(* IEC 61131-3 sources: plcassist-cli/packages/volt-lsp-iec/test-corpus/pro2193/Device/Plc Logic/Application/09 Misc/Library Manager/L_MC1P_MotionControlBasic (part 2) *)

(* ---- AXIS_REF.fb ---- *)
FUNCTION_BLOCK AXIS_REF EXTENDS L_DCO_AXIS_REF_BASE
VAR_INPUT
	LRVELOVERRIDE : LREAL := 1.0;
	LRACCOVERRIDE : LREAL := 1.0;
	LRJERKOVERRIDE : LREAL := 1.0;
	LRCOMMANDEDPOSITION : LREAL;
	LRCOMMANDEDVELOCITY : LREAL;
	LRCOMMANDEDACCELERATION : LREAL;
	LRSETVELOCITYLIMITHIGH : LREAL := 0;
	LRSETVELOCITYLIMITLOW : LREAL := 0;
	LRTORQUELIMHIGH : LREAL;
	LRTORQUELIMLOW : LREAL;
	LRTORQUELIMAUX : LREAL;
	SITORQUELIMDIR : SINT;
	XDELETETORQUELIM : BOOL;
	XSETTORQUELIMAUX : BOOL;
	XTORQUELIMHIGHFROMAPP : BOOL;
	XTORQUELIMLOWFROMAPP : BOOL;
	ITORQUELIMHIGHPCT : INT := 2000;
	ITORQUELIMLOWPCT : INT := 2000;
	EDIRECTION : MC_DIRECTION;
	XDRIVEENABLE : BOOL;
	XERRORRESET : BOOL;
	LRREFOFFSET : LREAL;
	LRREFOFFSETACT : LREAL;
	XENABLEPOSITIVE : BOOL := TRUE;
	XENABLENEGATIVE : BOOL := TRUE;
	LRSETSUPERACC : LREAL;
	LRSETSUPERVEL : LREAL;
	LRSETSUPERPOS : LREAL;
	LRSETMOVEACC : LREAL;
	LRSETMOVEVEL : LREAL;
	LRSETMOVEPOS : LREAL;
	XBUFCMDDONE : BOOL;
	XBUFRESTART : BOOL;
	LRPROFILESPEEDFIRST : LREAL;
	LRPROFILETARGETSPEED : LREAL;
	DWBUFFERCMD : __XWORD;
	XDISABLEERRORLOGGING : BOOL;
	XMOVEFUNBUSY : BOOL;
	XSUPERFUNBUSY : BOOL;
	LRCOMMANDEDPOSABSOLUT : LREAL;
	XRESETFOLLOWINGERROR : BOOL;
	XSETAXISQSP : BOOL;
	XSETDRIVEQSP : BOOL;
	EAXISSTATE : L_MC1P_AXIS_STATE := 2;
	LRSETPOSITION : LREAL := 0.0;
	LRSETVELOCITY : LREAL := 0.0;
	LRSETACCELERATION : LREAL := 0.0;
	LRSETTORQUE : LREAL := 0.0;
	LRVLTARGETVEL : LREAL := 0.0;
	LRLIMITEDVELOCITY : ARRAY [1..4] OF LREAL;
	LRLIMITEDDECTIME : ARRAY [1..4] OF LREAL;
	LRRESETSLSOFFSETVELOCITY : LREAL;
	DWLIMITERCONTROLACT : DWORD;
	SCSTOPAXISBYAPPL : L_MC1P_StopOperation;
	XSTAYINLASTSTATEREQUEST : BOOL;
	XMOVELASTSETPOSREQUEST : BOOL;
	LRSETVELMOVELASTSETPOS : LREAL;
	LRSETACCMOVELASTSETPOS : LREAL;
	LRSETDECMOVELASTSETPOS : LREAL;
	LRSETJERKMOVELASTSETPOS : LREAL;
	EDIRECTIONMOVELASTSETPOS : MC_DIRECTION;
	EDIRECTIONACTPROFILE : MC_DIRECTION;
	WAXISCONTROL : WORD := 0;
	XALLOWCHANGEOFCINHPAR : BOOL := FALSE;
	LRMOVEVELOFFSETVEL : LREAL;
	EOPTIMIZEDPROFILECALCULATIONMODE : UINT := 1;
	XLEAVESERVICESTATE : BOOL;
	XLEAVESERVICESTATEDISABLEDRIVE : BOOL;
	WLEAVESERVICESTATEPOWID : WORD;
END_VAR
VAR_OUTPUT
	EDEVICE : L_MC1P_DriveType := 0;
	WAXISSTATUS : DWORD := 0;
	EACTIVEERRORID : WORD := 0;
	LRACTPOSITION : LREAL := 0.0;
	LRACTVELOCITY : LREAL := 0.0;
	LRACTACCELERATION : LREAL := 0.0;
	LRACTTORQUE : LREAL := 0.0;
	LRSETTORQUETODRIVE : LREAL := 0;
	LRACTFOLLOWINGERROR : LREAL := 0.0;
	LRMAXFOLLOWINGERROR : LREAL := 0.0;
	XVIRTUAL : BOOL;
	XAXISAVAILABLE : BOOL;
	EACTDIRECTION : MC_DIRECTION;
	LRDIRECTIONHYSTERESISPOS : LREAL;
	LRDIRECTIONHYSTERESISTOL : LREAL := 1E-06;
	XDRIVEENABLED : BOOL;
	XERROR : BOOL;
	XWARNING : BOOL;
	XDRIVEERROR : BOOL;
	XDRIVEWARNING : BOOL;
	DWDRIVEERRORID : DWORD;
	XHOMEPOSAVAILABLE : BOOL;
	XSWLIMITENABLED : BOOL;
	XSWLIMITPOS : BOOL;
	XSWLIMITNEG : BOOL;
	XHWLIMITPOS : BOOL;
	XHWLIMITNEG : BOOL;
	XSPEEDEQZERO : BOOL;
	XINPOSITION : BOOL;
	LRTASKCYCLE : LREAL := 0.001;
	LRINVTASKCYCLE : LREAL := 1000.0;
	LRSWLIMITPOS : LREAL := 0.0;
	LRSWLIMITNEG : LREAL := 0.0;
	LRLASTSETPOSITION : LREAL;
	LRLASTTARGETPOSITION : LREAL;
	XSTANDSTILLSETVELOCITY : BOOL;
	XSTANDSTILLACTVELOCITY : BOOL;
	XSTOACTIVE : BOOL;
	XVOLTAGEENABLED : BOOL;
	XAXISREADYTOSWITCHON : BOOL;
	XAXISREADYFORMOTION : BOOL;
	SCPAR : L_MC1P_ParAccess;
END_VAR
VAR
	DWAXISCONFIGSETTINGS : DWORD;
	XSETVALUESAVAILABLE : BOOL;
	BYSETVALUESVALID : BYTE;
	DWTASKYCLE_US : DWORD := 1000;
	XSUSPENDFOLLOWINGERRORINT : BOOL;
	XSUSPENDFOLLOWINGERROREXT : BOOL;
	LRMAXVELOCITYAPPLOLD : LREAL;
	LRMAXACCELERATIONAPPLOLD : LREAL;
	LRMAXJERKAPPLOLD : LREAL;
	LRSWLIMITPOSOLD : LREAL;
	LRSWLIMITNEGOLD : LREAL;
	XENABLEPOSOLD : BOOL;
	XENABLENEGOLD : BOOL;
	DWLIMITERCONTROLOLD : DWORD;
	LRLIMITEDVELOCITYOLD : ARRAY [1..4] OF LREAL;
	LRLIMITEDDECTIMEOLD : ARRAY [1..4] OF LREAL;
	LRLIMITEDJERKOLD : ARRAY [1..4] OF LREAL;
	ELIMITERSTOPREACTION : L_IE1P_SeverityLevel := L_IE1P_SeverityLevel.WARNING;
	XSWLIMITDISABLE : BOOL := FALSE;
	XSWLIMITPOSNEU : BOOL;
	XSWLIMITPOSISTAN : BOOL;
	XSWLIMITNEGNEU : BOOL;
	XSWLIMITNEGISTAN : BOOL;
	PBYCOUPLEDMASTERAXIS : POINTER TO BYTE;
	PBYCOUPLEDPHASINGMASTERAXIS : POINTER TO BYTE;
	LRPHASESHIFTPOS : LREAL;
	LRPHASESHIFTVEL : LREAL;
	LRPHASESHIFTACC : LREAL;
	LRPHASESHIFTPOSOLD : LREAL;
	LRPHASESHIFTVELOLD : LREAL;
	LRPHASESHIFTACCOLD : LREAL;
	XSETPHASESHIFTVALUES : BOOL;
	ETRAVERSINGRANGEACT : L_MC1P_TraversingRange := 0;
	LRCYCLELENGTHACT : LREAL := 360.0;
	XENABLEHWLIMITPOS : BOOL := TRUE;
	XENABLEHWLIMITNEG : BOOL := TRUE;
	XHWSIGNALNEG : BOOL := FALSE;
	XHWSIGNALPOS : BOOL := FALSE;
	BHWENSCHPOSNEU : BOOL := TRUE;
	BNOTIFYERRORHWLIMITPOSISTAN : BOOL;
	BHWENSCHNEGNEU : BOOL := TRUE;
	BNOTIFYERRORHWLIMITNEGISTAN : BOOL;
	XAXISISHOMESOURCE : BOOL;
	XHOMEPOSAVAILABLEDRIVE : BOOL;
	SCHOMEPARAMETER : L_MC1P_HomeParameter;
	LRHOMEPOSITION : LREAL;
	XPOSCTRL : BOOL;
	XTPSUPPORTED : BOOL := FALSE;
	XTPWITHTIMESTAMP : BOOL := FALSE;
	SNTPMAXCHANNEL : SINT;
	PG : L_MC1P_PosProfiler := STRUCT(wCalcProfileMode := 1);
	ITFPG_MOVEACTIVE : L_MC1P_IPosProfilerActive;
	PG_MOVE : L_MC1P_PosProfiler := STRUCT(wCalcProfileMode := 1);
	ITFPG_SUPERACTIVE : L_MC1P_IPosProfilerActive;
	PG_SUPER : L_MC1P_PosProfiler := STRUCT(wCalcProfileMode := 1);
	PG_DUMMY : L_MC1P_PosProfiler := STRUCT(wCalcProfileMode := 1);
	SCPARAMSTOP : L_MC1P_ProfileParameter;
	XCTRLMODECHANGEREQ : BOOL;
	LRCTRLMODECHANGEREQACTVEL : LREAL;
	PFBMOVEBASIC : POINTER TO L_MC1P_MoveBasic;
	PFBMOVEBASICSUPER : POINTER TO L_MC1P_MoveBasic;
	XRESTARTPOSITIONING : BOOL;
	LRSETPOSITIONOLD : LREAL;
	LRSETVELOCITYOLD : LREAL;
	LRSETACCELERATIONOLD : LREAL;
	WACTFUNID : WORD := 0;
	WACTSUPERFUNID : WORD := 0;
	WACTPHASEFUNID : WORD := 0;
	PSERRORINST : POINTER TO STRING;
	SERRORINST : STRING;
	ERRORMANAGER : L_IE1P_ErrorManager;
	ERRORRESETOCCUREDTIMEWITHOUTLEM : SYSTIME;
	ASCERRORINFO : REFERENCE TO ARRAY [0..7] OF L_IE1P_ErrorInformation;
	ASCWARNINGINFO : REFERENCE TO ARRAY [0..7] OF L_IE1P_ErrorInformation;
	WINITSTATE : WORD;
	PAPPLICATION : POINTER TO APPLICATION;
	ATPDATA : ARRAY [1..4] OF L_MC1P_TPData;
	ATPDATASAVE : L_MC1P_TPData;
	XHOMINGSUPPORTED : BOOL;
	EAXISSTATEOLD : L_MC1P_AXIS_STATE := L_MC1P_AXIS_STATE.Disabled;
	ECONTROLMODE : L_MC1P_ControlMode := L_MC1P_ControlMode.PosCtrlDrive;
	ECONTROLMODEDEFAULT : L_MC1P_ControlMode := L_MC1P_ControlMode.PosCtrlDrive;
	ECONTROLMODEDEFAULTINT : L_MC1P_ControlMode := L_MC1P_ControlMode.PosCtrlDrive;
	POSCTRLDRIVEAVAILABLE : L_IE1P_Error;
	POSCTRLPLCAVAILABLE : L_IE1P_Error;
	SPEEDCTRLDRIVEAVAILABLE : L_IE1P_Error;
	TORQUECTRLDRIVE : L_IE1P_Error;
	XDRIVEENABLEOLD : BOOL;
	XLOCKEDFORSINGLEMOTION : BOOL := FALSE;
	XHOMEABSSWITCH : BOOL;
	XHOMEABSSWITCHOVERWRITEACTIVE : BOOL;
	XRAMPTOSTANDSTILL : BOOL;
	XRAMPTOSTANDSTILLDONE : BOOL;
	XRAMPTOSTANDSTILLACTIVE : BOOL;
	XDRIVEENABLEDOLD : BOOL;
	XDRIVEENABLEDREAL : BOOL;
	XDRIVEENABLEDREALOLD : BOOL;
	LRFOLLOWINGERRORINT : LREAL;
	XSUPPORTBRAKE : BOOL := FALSE;
	XSUPPORTDCBRAKE : BOOL := FALSE;
	XUSEASVIRTUALEXT : BOOL := FALSE;
	XUSEASVIRTUALEXTACT : BOOL := FALSE;
	LRSETSUPERACCOLD : LREAL;
	LRSETSUPERVELOLD : LREAL;
	LRSETSUPERPOSOLD : LREAL;
	ITFPARA : L_MC1P_IPara;
	XFASTSTOPDONE : BOOL;
	XFASTSTOPDONESAVE : BOOL;
	XSETFASTSTOPINT : BOOL;
	XERRRORSTOPACTIVE : BOOL;
	XERRRORSTOPDONE : BOOL;
	XSETAXISQSPACTIVE : BOOL;
	XRAMPQSPSTARTCALLEDFROMAPP : BOOL;
	XDRIVEQSPACTIVE : BOOL;
	XDRIVEQSPACTIVEOLD : BOOL;
	XDRIVEQSPSET : BOOL;
	XSETDRIVEFAILQSP : BOOL;
	XSETDRIVEFAILCINH : BOOL;
	XDRIVEQSPDONE : BOOL;
	XDRIVEQSPDONESAVE : BOOL;
	ESTOPTYPE : WORD;
	POW : L_MC1P_Power_Internal;
	XOBERVERESWITCHONTIME : BOOL := TRUE;
	FBBASE : L_MC1P_Template_ForAxis;
	ABC : L_MC1P_AxisBasicControl_Internal;
	ABCDATA : L_MC1P_AxisBasicControlInstanceData;
	ITFENCODER : L_MC1P_IEncoderInterface;
	ITFENCODERHANDLER : L_MC1P_IEncoderInterface;
	LRSETTORQUEFROMAXESGROUP : LREAL := 0;
	EPRECONTROLMODE : L_MC1P_PreControlMode := L_MC1P_PreControlMode.Automatic;
	GUID : L_MC1P_AxisGUID;
	LRTORQUEPRECTRL : LREAL;
	LRTORQUESET : LREAL;
	XMOVEFUNBUSYOLD : BOOL;
	XMOVEFUNBUSYOLDOLD : BOOL;
	DWIODRVDEVICEID : DWORD;
	WIODRVDEVICETYPE : WORD;
	EDEVICEORIGIN : L_MC1P_DriveType := L_MC1P_DriveType.Virtual;
	EDEVICECLASS : L_MC1P_DeviceClass := L_MC1P_DeviceClass.VirtualAxis;
	DWTARGETID : DWORD := 0;
	XCTRLFIRMWARECHECKPASSED : BOOL := FALSE;
	XENABLELOGENTRY : BOOL := 1;
	ETRAVERSINGRANGE : L_MC1P_TraversingRange := 1;
	LRCYCLELENGTH : LREAL := 360.0;
	LRINVCYCLELENGTH : LREAL := (1.0 / 360.0);
	LRDEFAULTVELOCITY : LREAL := 0.0;
	LRDEFAULTACCELERATION : LREAL := 0.0;
	LRDEFAULTJERK : LREAL := 0.0;
	LRMAXVELOCITYAPPL : LREAL := 0.0;
	LRMAXACCELERATIONAPPL : LREAL := 0.0;
	LRMAXJERKAPPL : LREAL := 0.0;
	XENABLESWLIMIT : BOOL := 0;
	WBEHAVEONSWLIMIT : WORD := 1;
	LRDECERRORSTOP : LREAL := 3600.0;
	LRJERKERRORSTOP : LREAL := 0.0;
	XREAKTONMCFBERROR : BOOL := 1;
	LRWINDOWSTANDSTILL : LREAL := 0.0;
	LRWINDOWVELOCITYCONST : LREAL := 0.0;
	LRWINDOWTARGETREACHED : LREAL := 0.0;
	LRWINDOWTARGETREACHEDTIME : LREAL := 0.0;
	LRMODPOSTOLERANCE : LREAL := 0.0;
	XSETVALUEMONITORING : BOOL := 0;
	EPARAMETERINDEX : WORD := 101;
	DWPARABASEINDEX : DWORD;
	PPARA2 : L_SSYP.L_SSYP_EVTPARAM_CmpLenzeIPCSystemSoftPLCParaChanged;
	HEVENTPARWRITE : SysTypes.RTS_IEC_HANDLE;
	HINTERFACEPARWRITE : SysTypes.RTS_IEC_HANDLE;
	HEVENTDOWNLOADDONE : SysTypes.RTS_IEC_HANDLE;
	HINTERFACEDOWNLOADDONE : SysTypes.RTS_IEC_HANDLE;
	HEVENTRESETDONE : SysTypes.RTS_IEC_HANDLE;
	HINTERFACERESETDONE : SysTypes.RTS_IEC_HANDLE;
	ITFCALLBACK : CmpEventMgr.ICmpEventCallback;
	DWEVENTCOUNTER : DWORD;
	WENABLEDRIVEBLOCKEDBYOBJECTTRANSFER : WORD := 0;
	XUSEDBYAXESGROUP : BOOL;
	PUSEDAXESGROUP : POINTER TO BYTE;
	DWEVTINITCOUNT : DWORD;
	XNEWHOMEPOSLOADED : BOOL;
	DWSETPOSITIONCALLCYCLE : DWORD;
	XSETPOSITIONCALLCYCLEVALID : BOOL;
	AITFFILTER : ARRAY [1..c_MaxFilterInt] OF L_MC1P_ISetvalueManipulationInterface;
	XENABLEFILTER : BOOL;
	XFILTERAVAILABLE : BOOL;
	XIGNORFILTERINSTOP : BOOL := TRUE;
	XIGNORFILTERINSTOPITF : BOOL;
	XUSEFILTERVALUESFORSYNC : BOOL := FALSE;
	LRSETPOSITIONFILT : LREAL;
	LRSETVELOCITYFILT : LREAL;
	LRSETACCELERATIONFILT : LREAL;
	LRSETTORQUEFILT : LREAL;
	LRSETVALUEFILTERPOSDEVIATION : LREAL;
	XINTARGETSETVALUEFILTER : BOOL;
	XSUSPENDSETVALUEFILTERCALL : BOOL := FALSE;
	LRSETPOSITIONFILTOLD : LREAL;
	LRSETVELOCITYFILTOLD : LREAL;
	LRSETACCELERATIONFILTOLD : LREAL;
	LRSETTORQUEFILTOLD : LREAL;
	LRSETPOSROUNDSFILTOLD : LREAL;
	AITFCOMPENSATION : ARRAY [1..c_MaxFilterInt] OF L_MC1P_ICompensationInterface;
	LRCOMPENSATIONOFFSETPOS : LREAL;
	LRCOMPENSATIONOFFSETVEL : LREAL;
	LRCOMPENSATIONOFFSETACC : LREAL;
	LRACTPOSITIONUNFILTERED : LREAL;
	LRINTARGETPOS : LREAL;
	LRACTTIMETARGETREACHED : LREAL;
	XSETVALUEINTARGET : BOOL;
	XUSEACYCLIC : BOOL := FALSE;
	XFORCEACYCLICMODE : BOOL := FALSE;
	WAXISMODE : WORD := 1;
	WAXISMODEOLD : WORD := 255;
	LRTRANSMITCYCLESACTPOS : LREAL := 0.0;
	LRTRANSMITCYCLESSETPOS : LREAL := 1.0;
	XCONNECTORDISABLEDBYPROJECT : BOOL;
	XCONNECTORDISABLED : BOOL;
	XAXISDETECTIONBUSY : BOOL;
	XAXISDETECTED : BOOL;
	XCONFIGDONE : BOOL;
	XBASICINIT : BOOL := TRUE;
	XAXISCONNECTBUSY : BOOL;
	XAXISCONNECTDONE : BOOL;
	XPDOINTERFACEDISABLED : BOOL;
	XDRIVETESTMODEACTIVE : BOOL;
	LRACTPOSROUNDS : LREAL;
	LRSETPOSROUNDS : LREAL;
	LRSETPOSROUNDSFILT : LREAL;
	LRSETPOSROUNDSLAST : LREAL;
	LRTARGETPOSROUNDS : LREAL;
	XTARGETPOSVALID : BOOL;
	XTARGETPOSFROMMOVEREL : BOOL;
	LISETPOSCYCLE : LINT;
	LISETPOSCYCLERES : UDINT;
	XSETPOSCYCLEZERO : BOOL;
	XRECOVERLASTSETPOS_RAMP : BOOL := FALSE;
	XRECOVERLASTSETPOS_POSCTRL : BOOL := TRUE;
	XRECOVERYPOSVALID : BOOL;
	XMOVELASTSETPOS : BOOL;
	LRRECOVERYWINDOWPOS : LREAL;
	LRRECOVERYWINDOWNEG : LREAL;
	LRRECOVERYPOSITION : LREAL;
	LRRECOVERYVEL : LREAL := 360;
	LRRECOVERYACC : LREAL := 3600;
	LRRECOVERYDEC : LREAL := 3600;
	LRRECOVERYJERK : LREAL := 0;
	XSLSACTIVE : BOOL;
	XSLSACTIVEOLD : BOOL;
	XSLIREQUESTACTIVE : BOOL;
	XSWLIMITSACTIVE : BOOL;
	LRSLIDISTANCE : LREAL := 360;
	LRSLSVELOCITY : LREAL;
	LRSLSVELOCITYOLD : LREAL;
	LRSLSDECELERATION : LREAL;
	LRSLSDECELERATION2 : LREAL;
	LRSLSDECELERATIONOLD : LREAL;
	LRSLSJERK : LREAL;
	XSLSCHANGES : BOOL;
	XSLSNEWACTIVEDECELERATION : BOOL;
	WSLSWARNING : WORD;
	XLIMITERENABLEPOSITIVE : BOOL := TRUE;
	XLIMITERENABLENEGATIVE : BOOL := TRUE;
	XLIMITERENABLED : BOOL;
	XLIMITATIONSLSACTIVE : BOOL;
	XLIMITATIONACTIVE : BOOL;
	LRSLSDECTIME : LREAL := 100;
	LRSLSDECTIMEOLD : LREAL := 100;
	WSAFESTOPCONTROLWORD : WORD;
	WSAFESTOPCONTROLWORDOLD : WORD;
	READPARAMETER : L_DCO_ReadDriveParameter;
	WRITEPARAMETER : L_DCO_WriteDriveParameter;
	DWACTUALSPEEDCONTROLLERLIMIT : DWORD;
	XLIMITSPEEDCONTROLLERSLS : BOOL;
	DWDISABLESAFETYINTERFACE : DWORD;
	DWREQUESTSAFETYINTERFACE : DWORD;
	XFOLLOWERSLS : BOOL;
	LRSLSTIMER : LREAL;
	LRSLSTIMERTEMP : LREAL;
	XSLSACTIVATED : BOOL := FALSE;
	XSETSTOPBYDIRECTIONACTIVE : BOOL;
	XSETSTOPBYLIMITERACTIVE : BOOL;
	XSETSTOPCINHBYLIMITERACTIVE : BOOL;
	XSLSVELOCITYACTIVE : BOOL;
	XSLSDECTIMEACTIVE : BOOL;
	XSLSWARNINGACTIVE : BOOL;
	ETYPEFUNCTIONACT : L_MC1P_TypeFunction := L_MC1P_TypeFunction.Type_Any;
	SCSTOPBYERROR : L_MC1P_StopOperation;
	SCSTOPBYAXESGROUP : L_MC1P_StopOperation;
	DWAXISERRORITFID : DWORD := 0;
	ICMODE : WORD;
	ICMODEOLD : WORD;
	DWIC : DWORD;
	DWICOLD : DWORD;
	XINTERNALCONTROLMODEACTIVE : BOOL;
	XINTERNALCONTROLMODEACTIVEOLD : BOOL;
	XREFDUMMY : BOOL;
	LRREFDUMMY : LREAL;
	RREFDUMMY : REAL;
	WREFDUMMY : WORD;
	IREFDUMMY : INT;
	DWREFDUMMY : DWORD;
	DIREFDUMMY : DINT;
	LWREFDUMMY : LWORD;
	LIREFDUMMY : LINT;
	SREFDUMMY : STRING;
	USIREFDUMMY : USINT;
	BYREFDUMMY : BYTE;
	UIREFDUMMY : UINT;
	UDIREFDUMMY : UDINT;
	ULIREFDUMMY : ULINT;
	DWCALLCYCLE : DWORD;
	DWCALLCYCLE_US : DWORD;
	DWTPDELAYACTPOS : DWORD := 0;
	DWACTDCTIME : DWORD;
	PDWABSOLUTECOUNTER : POINTER TO DWORD;
	XGLOBALTIMESTAMPSUPPORTED : BOOL;
	HMOTIONTASK : SysTypes.RTS_IEC_HANDLE := 0;
	WACTPOSIDX : WORD;
	ADWACTTIMESTAMPS : ARRAY [0..15] OF DWORD;
	ALRACTPOSITION : ARRAY [0..15] OF LREAL;
	ALRACTPOSITIONUNFILTERED : ARRAY [0..15] OF LREAL;
	ALRACTPOSROUNDS : ARRAY [0..15] OF LREAL;
	ALRTPPOSOFFSET : ARRAY [0..15] OF LREAL;
	HEVENTRESETOCCURED : SysTypes.RTS_IEC_HANDLE := SysTypes.RTS_INVALID_HANDLE;
	HINTERFACERESETOCCURED : SysTypes.RTS_IEC_HANDLE := SysTypes.RTS_INVALID_HANDLE;
	XGENERRORREAKTINDEVICE : BOOL;
	XFORWARDERRORSASWARNINGS : BOOL;
	WEVTCOUNT_SETERRORREACTION : WORD;
	WEVTCOUNT_UPDATEACTIVEERROR : WORD;
	WEVTCOUNT_RESETOCCURED : WORD;
	XINTERNALERRORRESET : BOOL;
	XINTERNALERRORRESETFROMLEM : BOOL;
	WHANDLINGLEM : WORD := 0;
	XERRORRESETREQUESTSEND : BOOL;
	WERRORRESETREQUESTSEND : WORD := 0;
	RESETINTERNAL : L_MC1P_Reset_Internal;
	DWACTSTATEDETERMINEEVENT : DWORD;
	SEVERITYCMDEXT : USINT;
	EERRORREACTIONCMDEXT : L_IE1P_SeverityLevel := L_IE1P_SeverityLevel.NO_RESPONSE;
	DWERRORINFOEXT : DWORD;
	XEXTERROR : BOOL;
	MYSYSTEMSEVERITY : USINT;
	XJOGGINGACTIVE : BOOL;
	LRJOGGINGSETVEL : LREAL := 360.0;
	LRJOGGINGSETACC : LREAL := 360.0;
	LRJOGGINGSETDEC : LREAL := 1440.0;
	LRJOGGINGSETJERK : LREAL := 0.0;
	XJOGUSEAXISPAR : BOOL := FALSE;
	XHOMEPOSUSEAXISPAR : BOOL := FALSE;
	XUSEFASTSTOPBEHAVIOUR : BOOL := TRUE;
	XFIRSTBASEINITDONE : BOOL := FALSE;
	EHWLIMITERRORREACTION : USINT := 19;
	ESWLIMITERRORREACTION : USINT := 19;
	ELIMITPROFILEERRORREACTION : USINT := 2;
	ECINHERRORREACTION : USINT := 19;
	LRREFROUNDS : LREAL;
	XMOVELASTSETPOSACTIVE : BOOL;
	XSTAYINLASTSTATEACTIVE : BOOL;
	XABORTSTAYINLASTSTATEREQUEST : BOOL;
	XCINHACTIVE : BOOL;
	XCINHACTIVEOLD : BOOL;
	XSTOACTIVEOLD : BOOL;
	XSETPOSINSIDEWINDOW : BOOL;
	XSTAYINLASTSTATEACTIVEOLD : BOOL;
	XDRIVESTATEBEFORECINH : BOOL;
	LRPOSOFFSETMOVELASTSETPOS : LREAL;
	LRVELOFFSETMOVELASTSETPOS : LREAL;
	LRACCOFFSETMOVELASTSETPOS : LREAL;
	XHALTPARAMETERSUPPORTED : BOOL;
	LRHALTDEC : LREAL := 1800;
	LRHALTJERK : LREAL := 0;
	XHALTBYABC : BOOL;
	SCTIMESTAMP : L_MC1P_TimeStamp;
	XACTIVATETIMEMEASUREMENT : BOOL;
	XISSAFETYDEVICE : BOOL;
	WINDEXINT : WORD;
	BYSUBINDEXINT : BYTE;
	BYSLSREADWRITECOUNTER : BYTE;
	XCALCMODULOASLIMITED : BOOL := FALSE;
	FBSTEADYSTATE : L_MC1P_SteadyState;
	WDEVICETYPETEMP : WORD;
	DWIODRVDEVICEIDTEMP : DWORD;
	XUSEQSPDRIVEINSTEADOFQSPAPPL : BOOL := FALSE;
	XMINJERKAVAILABLE : BOOL;
	XMINJERKAVAILABLEOLD : BOOL;
	XMINJERKACTIVE : BOOL;
	XMINJERKACTIVEOLD : BOOL;
	LRMINJERK : LREAL;
	LRMINJERKOLD : LREAL;
	LRMOVEVELOFFSETVELOLD : LREAL;
	XSETVALUESFORINTERNALSTOPAVAILABLE : BOOL;
	XSETVALUESFROMINTERNALSTOPACTIVE : BOOL;
	XOPTRAMPSFORMANUALJOG : BOOL := TRUE;
	XCHANGECINHPARNOTALLOWED : BOOL := FALSE;
	XBEHAVIOURFORVIRTUALMASTER : BOOL := FALSE;
	STOPAXISBYERRORREACTIONCOUNTER : L_IE1P_ReactionCounter;
	SCSTOPAXISBYERRORREACTION : L_MC1P_StopOperation;
	MODULEHANDLERBASE : L_IMHP_ModuleHandler := STRUCT(CompActiveDefault := FALSE, Layer := L_IMHP_Layer.Motion, CompType := L_IMHP_ComponentType.VirtualAxis);
	FB_GETDIRECTIONACTVALUES : L_MC1P_GetDirection;
	WDIRECTIONSETVALUES : WORD;
	XQSPWITHOUTREACTION : BOOL;
	XVALIDMFEFWVERSION : BOOL;
	XSETDRIVEQSPDISABLED : BOOL;
	EKINDOFMOTIONSELECTION : L_MC1P_KindOfMotion;
	EACTIVEUNIT : WORD;
	WERRORIDINITSTATE : WORD;
	ITFMANIPULATEACTVALUES : L_Mc1P_IManipulateActValues;
	XSETVELOCITYGTSLS : BOOL;
	XCLOSEBRAKEATQSPRAMPEND : BOOL;
	C_STRNOERROR : STRING := '-';
	C_STRUNDEFERROR : STRING := 'undefined';
	C_MAXFILTER : WORD := 2;
	C_MAXCOMP : WORD := 2;
	C_MAXFILTERINT : WORD := (c_MaxFilter + 1);
	C_UDILOGCOMPONENDID : UDINT := 16#2800;
	ACTACCELERATION : LREAL;
	ACTPOSITION : LREAL;
	ACTTORQUE : LREAL;
	ACTVELOCITY : LREAL;
	AXISPOOLCOUNT : WORD;
	AXISSLOT : L_MC1P_AxisSlot;
	CIA402ADVANCEDAXIS : BOOL;
	CMDCINH : BOOL;
	CMDFASTSTOP : BOOL;
	CMDFASTSTOPCINH : BOOL;
	CMDQSP : BOOL;
	CMDQSPCINH : BOOL;
	CYCLELENGTH : LREAL;
	FEEDCONSTANT : LREAL;
	GETACTIVELIMTERCONTROLWORD : DWORD;
	GETMASTERID : POINTER TO BYTE;
	HOMEPOSPERMANTENTSETACTIVE : BOOL;
	HOMEPOSPERMANTENTSETACTIVELOADENCODER : BOOL;
	LICENSECONFIG : STRING;
	MODULEHANDLER : L_IMHP_IModuleHandler;
	QSPATFASTSTOPEND : BOOL;
	QSPWITHOUTREACTION : BOOL;
	RESETFOLLOWINGERRORATFASTSTOPEND : BOOL;
	SERVICEDIRECTION : L_MC1P_ServiceDirection;
	SETACCELERATIONFORSYNC : LREAL;
	SETHOMEPOSSTATEINDEPENDENTACTIVE : BOOL;
	SETPOSITIONFORSYNC : LREAL;
	SETPOSROUNDS : LREAL;
	SETTORQUEFORSYNC : LREAL;
	SETVELOCITYFORSYNC : LREAL;
	STARTPOSFORINTERNALSTOP : LREAL;
	TASKCYCLE : LREAL;
	TIMEDELAYACTPOS : LREAL;
	TIMEDELAYSETPOS : LREAL;
	TRAVERSINGRANGE : L_MC1P_TraversingRange;
	USEDASINTERNALAXISINSTANCE : BOOL;
	USEDBYVIRTUALMASTER : BOOL;
END_VAR
END_FUNCTION_BLOCK

METHOD ACTIVATEACYCLICMODE
VAR_INPUT
	XACTIVATE : BOOL;
END_VAR
END_METHOD

METHOD CALCACTDIRECTION
END_METHOD

METHOD CALCACTPOSUNFILTERED : LREAL
END_METHOD

METHOD CALCSETDIRECTION : WORD
VAR_INPUT
	LRCYCVELIN : LREAL;
END_VAR
END_METHOD

METHOD CALLSIMULATION
VAR_INPUT
	CALLSTATE : L_UBUP_StateHandleCase;
END_VAR
END_METHOD

METHOD CHECKDIRECTION : BOOL
VAR_INPUT
	DIRECTION : MC_DIRECTION;
	ETYPEFUNCTION : L_MC1P_TypeFunction;
END_VAR
END_METHOD

METHOD CHECKMAXMODULOPOSDIFF
END_METHOD

METHOD CHECKPLNOTVALID : BOOL
END_METHOD

METHOD CHECKPLAUSIBILITYOFSETVALUES
END_METHOD

METHOD CHECKPOWER : BOOL
VAR_INPUT
	DWPOSSTATE : DWORD;
	LRVEL : LREAL;
END_VAR
END_METHOD

METHOD CHECKSLSVELOCITY : BOOL
END_METHOD

METHOD CHECKSETPOSINWINDOW : BOOL
END_METHOD

METHOD COMPENSATELOADPOSOFFSET
END_METHOD

METHOD ENABLEDRIVE : BOOL
VAR_INPUT
	XENABLE : BOOL;
END_VAR
END_METHOD

METHOD FLOATTOFRAC
VAR_INPUT
	LRINPUT : LREAL;
	PDIINTEGER : POINTER TO DINT;
	PUDIRESIDUAL : POINTER TO UDINT;
END_VAR
END_METHOD

METHOD FLOATTOFRACLINT
VAR_INPUT
	LRINPUT : LREAL;
	PLIINTEGER : POINTER TO LINT;
	PUDIRESIDUAL : POINTER TO UDINT;
END_VAR
END_METHOD

METHOD GENACTVALUES
END_METHOD

METHOD GETACTVEL : LREAL
END_METHOD

METHOD GETACTVELOCITYEXACT : LREAL
END_METHOD

METHOD GETACTIVEQUICKSTOPOPTION : L_MC1P_QuickStopOption
END_METHOD

METHOD GETAXISSLOT : UINT
END_METHOD

METHOD GETBRAKE : POINTER TO L_MC1P_BrakeControlBase
END_METHOD

METHOD GETBRAKESERVICE : POINTER TO L_MC1P_BrakeService
END_METHOD

METHOD GETCOUPLEDMASTERAXIS : POINTER TO BYTE
END_METHOD

METHOD GETCOUPLEDPHASINGMASTERAXIS : POINTER TO BYTE
END_METHOD

METHOD GETDRIVESTATE : BOOL
END_METHOD

METHOD GETEFFECTIVEMFESPEEDOFFSET : INT
VAR_INPUT
	INOFFSET : INT;
END_VAR
END_METHOD

METHOD GETMODULODIFF : LREAL
VAR_INPUT
	LRDIFF : LREAL;
END_VAR
VAR_IN_OUT
	AXIS : AXIS_REF;
END_VAR
END_METHOD

METHOD GETMODULOPOSITION : LREAL
VAR_INPUT
	LRNEWPOS : LREAL;
END_VAR
VAR_OUTPUT
	LRROUNDS : LREAL;
END_VAR
VAR_IN_OUT
	AXIS : AXIS_REF;
END_VAR
END_METHOD

METHOD GETPGMOVE : REFERENCE TO L_MC1P_PosProfiler
VAR_INPUT
	ITFPGACTIVE : L_MC1P_IPosProfilerActive;
END_VAR
END_METHOD

METHOD GETPGDUMMY : REFERENCE TO L_MC1P_PosProfiler
END_METHOD

METHOD GETPGSUPER : REFERENCE TO L_MC1P_PosProfiler
VAR_INPUT
	ITFPGACTIVE : L_MC1P_IPosProfilerActive;
END_VAR
END_METHOD

METHOD GETPHASESHIFT
VAR_OUTPUT
	LRPOS : LREAL;
	LRVEL : LREAL;
	LRACC : LREAL;
END_VAR
END_METHOD

METHOD GETRECEIVEDATA : DWORD
VAR_INPUT
	LWMASK : LWORD;
END_VAR
END_METHOD

METHOD GETTPWITHPOSITIONACTIVE : BOOL
VAR_INPUT
	SITPNUMBER : SINT;
END_VAR
END_METHOD

METHOD GETTPWITHTIMESTAMPACTIVE : BOOL
VAR_INPUT
	SITPNUMBER : SINT;
END_VAR
END_METHOD

METHOD HALTCALLEDBYABC
VAR_INPUT
	XCALLEDBYABC : BOOL;
END_VAR
END_METHOD

METHOD HLP_MODULOPOS : LREAL
VAR_INPUT
	LRPOSITION : LREAL;
	LRCYCLELENGTH : LREAL;
END_VAR
END_METHOD

METHOD HLP_MODULOPOS2 : LREAL
VAR_INPUT
	LRPOSITION : LREAL;
	LRCYCLELENGTH : LREAL;
	LRINVCYCLELENGTH : LREAL;
END_VAR
END_METHOD

METHOD INTOLERANCEWINDOW : BOOL
VAR_INPUT
	LRPOSITION : LREAL;
END_VAR
VAR_OUTPUT
	DIRECTION : MC_DIRECTION;
END_VAR
END_METHOD

METHOD INTERNALCONTROLMODE
END_METHOD

METHOD ISINCLUDEDINRECEIVEDATA : BOOL
VAR_INPUT
	LWMASK : LWORD;
END_VAR
END_METHOD

METHOD ISINCLUDEDINTRANSMITDATA : BOOL
VAR_INPUT
	LWMASK : LWORD;
END_VAR
END_METHOD

METHOD ISMOTIONALLOWED : BOOL
VAR_INPUT
	ETYPEFUNCTION : L_MC1P_TypeFunction;
END_VAR
VAR_IN_OUT
	XSUPERIMPOSED : BOOL;
END_VAR
END_METHOD

METHOD ISMOTIONALLOWED2 : BOOL
VAR_INPUT
	ETYPEFUNCTION : L_MC1P_TypeFunction;
	XCHECKHOMEPOS : BOOL;
END_VAR
VAR_OUTPUT
	EERRORCAUSE : L_IE1P_Error := L_IE1P_Error.NoError;
END_VAR
VAR_IN_OUT
	XSUPERIMPOSED : BOOL;
END_VAR
END_METHOD

METHOD LEAVESERVICESTATE
END_METHOD

METHOD LEAVESERVICESTATEBEAVIOUR : DINT
VAR_INPUT
	XDISABLEDRIVE : BOOL;
END_VAR
END_METHOD

METHOD LEAVESERVICESTATESTART : BOOL
END_METHOD

METHOD LIMITPROFILEDATA : WORD
VAR_INPUT
	PPROFLE : POINTER TO L_MC1P_ProfileParameter;
	PPROFLEOLD : POINTER TO L_MC1P_ProfileParameter;
END_VAR
END_METHOD

METHOD LOCKEDFORSINGLEMOTION
VAR_INPUT
	XLOCKED : BOOL;
END_VAR
END_METHOD

METHOD REGISTERAXESGROUP : BOOL
VAR_INPUT
	XUNREGISTER : BOOL;
	PAXESGROUP : POINTER TO BYTE;
END_VAR
END_METHOD

METHOD REGISTERFUNCTION : WORD
END_METHOD

METHOD REGISTERPHASINGFUNCTION : WORD
VAR_INPUT
	PMASTERAXIS : POINTER TO BYTE;
END_VAR
END_METHOD

METHOD REGISTERSUPERFUNCTION : WORD
END_METHOD

METHOD REGISTERSYNCFUNCTION : WORD
VAR_INPUT
	PMASTERAXIS : POINTER TO BYTE;
END_VAR
END_METHOD

METHOD RESETERRORSTATEOFCOMMANDS : BOOL
END_METHOD

METHOD RESETFOLLOWINGERROR
END_METHOD

METHOD RESETMOVEBUFFEREDINFO
END_METHOD

METHOD RESETMOVEINFO
END_METHOD

METHOD SERVICEMODEHANDLINGINDRIVEACTIVE : BOOL
END_METHOD

METHOD SETACTPOSITION
VAR_INPUT
	POSITION : LREAL;
	RELATIVE : BOOL;
END_VAR
END_METHOD

METHOD SETAXISSTATUSWORD
END_METHOD

METHOD SETBUFFERDATAALLOWED : BOOL
VAR_INPUT
	EMODE : MC_BUFFER_MODE;
	LRSPEED1 : LREAL;
	LRSPEED2 : LREAL;
	DWINSTANCE : __XWORD;
END_VAR
END_METHOD

METHOD SETDCBRAKE
VAR_INPUT
	XSETDCBRAKE : BOOL;
END_VAR
VAR_OUTPUT
	XDCBRAKEACTIVE : BOOL;
END_VAR
END_METHOD

METHOD SETENCODERITF
VAR_INPUT
	ENCODERIN : L_MC1P_IEncoderInterface;
END_VAR
END_METHOD

METHOD SETHOMEABSSWITCH
VAR_INPUT
	HOMEABSSWITCH : BOOL;
END_VAR
END_METHOD

METHOD SETHOMEABSSWITCHOVERWRITE
VAR_INPUT
	XHOMEABSSWITCHSIGNAL : BOOL;
	XOVERWRITESIGNAL : BOOL;
END_VAR
END_METHOD

METHOD SETMACHINEDATA
END_METHOD

METHOD SETPHASESHIFT
VAR_INPUT
	LRPOS : LREAL;
	LRVEL : LREAL;
	LRACC : LREAL;
END_VAR
END_METHOD

METHOD SETPOSEQACTPOS
END_METHOD

METHOD SETPRECONTROLMODE
VAR_INPUT
	EPRECONTROLMODENEW : L_MC1P_PreControlMode := L_MC1P_PreControlMode.Automatic;
END_VAR
END_METHOD

METHOD SETTARGETPOS
VAR_INPUT
	LRTARGETPOSNEW : LREAL;
	LRTARGETPOSROUNDSNEW : LREAL;
	XVALID : BOOL;
END_VAR
END_METHOD

METHOD SETTARGETPOS2
VAR_INPUT
	LRTARGETPOSNEW : LREAL;
	LRTARGETPOSROUNDSNEW : LREAL;
	XVALID : BOOL;
	XRELMODE : BOOL;
END_VAR
END_METHOD

METHOD SETTORQUEVALUE
VAR_INPUT
	LRTORQUE : LREAL;
	WMODE : WORD;
END_VAR
END_METHOD

METHOD SETVELEQREFVALUE
VAR_INPUT
	LRREFVELOCITY : LREAL;
END_VAR
END_METHOD

METHOD SETVELOCITYOFFSET
VAR_INPUT
	WMODE : WORD;
	LROFFSETVELOCITY : LREAL;
END_VAR
END_METHOD

METHOD SPEEDEQZERO : BOOL
VAR_INPUT
	LRSPEEDIN : LREAL;
END_VAR
END_METHOD

METHOD SUSPENDFOLLOWINGERROR
VAR_INPUT
	XSUSPEND : BOOL;
END_VAR
END_METHOD

METHOD UPDATEERRORINFO
END_METHOD

METHOD UPDATEREADYFORMOTIONSTATUS : BOOL
VAR_INPUT
	AXISENABLED : BOOL;
END_VAR
END_METHOD

METHOD CALLRECIEVEPARAMETER
END_METHOD

METHOD CALLSDODATAHANDLING
END_METHOD

METHOD CALLTRANSMITPARAMETER
END_METHOD

METHOD CHECKCOMMUNCATION
END_METHOD

METHOD CHECKMAPPEDDATAVALID : BOOL
VAR_INPUT
	PADDDATA : POINTER TO BYTE;
	PDATA : POINTER TO POINTER TO BYTE;
END_VAR
VAR_OUTPUT
	XERROR : BOOL;
	EERRORID : L_IE1P_Error;
END_VAR
END_METHOD

METHOD GETMAPPEDDATA : POINTER TO BYTE
VAR_INPUT
	UIINDEX : WORD;
	USISUBINDEX : USINT;
	USISIZE : USINT;
	XWRITEACCESS : BOOL;
	PADDDATA : POINTER TO BYTE;
	PXWAITFORINITACCESS : POINTER TO BOOL;
END_VAR
VAR_OUTPUT
	EERRORID : L_IE1P_Error;
	XERROR : BOOL;
	USISIZEACT : USINT := 0;
END_VAR
END_METHOD

METHOD GETMAPPEDDATASUPPORT : BOOL
END_METHOD

METHOD RESETMAPPEDDATA
VAR_INPUT
	PADDDATA : POINTER TO BYTE;
END_VAR
END_METHOD

METHOD RESETSDODATA : DINT
VAR_INPUT
	IDX : DWORD;
	PDWSEMAPARACCESS : POINTER TO DWORD;
END_VAR
VAR_IN_OUT
	SDODATA : L_DCO_SdoData;
END_VAR
END_METHOD

METHOD CONFIGUREAXIS
END_METHOD

METHOD CONFIGUREAXIS2
END_METHOD

METHOD CONFIGUREAXISCONNECTOR
END_METHOD

METHOD CONFIGUREAXISCONNECTORBASICS : BOOL
END_METHOD

METHOD CONNECTCMDITFAUTOTUNING
END_METHOD

METHOD DETERMINETASKCYCLEINTERVAL : UDINT
END_METHOD

METHOD ENABLEAXISCONNECTOR : BOOL
END_METHOD

METHOD FINDANDCONNECTMOTIONUTILS
END_METHOD

METHOD GETTRANSMITCYCLESACTPOSFORPOSCTRL : LREAL
END_METHOD

METHOD REGISTERAXISPROPERTIES
END_METHOD

METHOD RESETAXISCONNECTOR
END_METHOD

METHOD SETAXISPROPERTIES
VAR_INPUT
	XUSEVIRTUAL : BOOL;
END_VAR
END_METHOD

METHOD UPDATEFATHERCONNECTOR
END_METHOD

METHOD CHECKAVAILABLECONTROLMODE : BOOL
END_METHOD

METHOD CONFIGURECONTROLMODE
VAR_OUTPUT
	EERRORID : L_IE1P_Error;
END_VAR
END_METHOD

METHOD GETDEFAULTCONTROLMODE : L_MC1P_ControlMode
END_METHOD

METHOD ISAVAILABLECONTROLMODE : BOOL
VAR_INPUT
	ECONTROLMODE : L_MC1P_ControlMode;
END_VAR
VAR_OUTPUT
	EERRORID : L_IE1P_Error;
END_VAR
END_METHOD

METHOD SETCONTROLMODE : BOOL
VAR_INPUT
	ECONTROLMODE : L_MC1P_ControlMode := L_MC1P_ControlMode.PosCtrlDrive;
	XKEEPACTPOSPRIORFDB : BOOL := FALSE;
	XRESTARTPOSITIONING : BOOL := FALSE;
END_VAR
VAR_OUTPUT
	EERRORID : L_IE1P_Error;
END_VAR
END_METHOD

METHOD SETCONTROLERITF
VAR_INPUT
	ITFCONTROLERNEW : L_MC1P_IControllerInterface;
END_VAR
END_METHOD

METHOD SETDEFAULTCONTROLMODE : BOOL
END_METHOD

METHOD CLEARERROR
VAR_INPUT
	PINSTANCE : POINTER TO BYTE := 0;
END_VAR
END_METHOD

METHOD CLEARERROR2
VAR_INPUT
	INSTANCEID : DWORD := 0;
END_VAR
END_METHOD

METHOD CLEARERRORID
VAR_INPUT
	PINSTANCE : POINTER TO BYTE := 0;
	WERRORID : WORD;
END_VAR
END_METHOD

METHOD CLEARERRORID2
VAR_INPUT
	INSTANCEID : DWORD := 0;
	WERRORID : WORD;
END_VAR
END_METHOD

METHOD CLEARERRORID3
VAR_INPUT
	INSTANCEID : DWORD := 0;
	WERRORID : WORD;
	DWEXTENDEDERRORINFO : DWORD;
END_VAR
END_METHOD

METHOD GETERRORITFID : DWORD
END_METHOD

METHOD HANDLEERRORENTRY : BOOL
VAR_INPUT
	WERRORID : L_IE1P_Error := 0;
	INSTANCEID : DWORD := 0;
	PSINSTANCENAME : POINTER TO BYTE := 0;
	DWEXTENDEDERRORINFO : DWORD;
	EERRORREACTION : L_IE1P_SeverityLevel := 0;
	XAUTORESET : BOOL;
	XNOLOGGINGENTRY : BOOL;
	XEXTERNALERROR : BOOL;
END_VAR
END_METHOD

METHOD NOTIFYERROR : BOOL
VAR_INPUT
	WERRORID : L_IE1P_Error := 0;
	PINSTANCE : POINTER TO BYTE := 0;
	PSINSTANCENAME : POINTER TO BYTE := 0;
	XSETERRORSTOP : BOOL := FALSE;
END_VAR
END_METHOD

METHOD NOTIFYERROR2 : BOOL
VAR_INPUT
	WERRORID : L_IE1P_Error := 0;
	INSTANCEID : DWORD := 0;
	PSINSTANCENAME : POINTER TO BYTE := 0;
	EERRORREACTION : L_IE1P_SeverityLevel := 0;
END_VAR
END_METHOD

METHOD SERERRORREACTIONEXTERN
VAR_INPUT
	EERRORREACTION : L_IE1P_SeverityLevel;
	WERRORID : WORD;
	INSTANCEID : DWORD := 0;
	XAUTORESET : BOOL;
	DWEXTENDEDERRORINFO : DWORD;
	XEXTERNALERROR : BOOL;
END_VAR
END_METHOD

METHOD UPDATEERRORREAKTION
VAR_INPUT
	SEVERITY : L_IE1P_SeverityLevel;
END_VAR
END_METHOD

METHOD EVENTCALLBACK : UDINT
VAR_INPUT
	PEVENTPARAM : POINTER TO EventParam;
END_VAR
END_METHOD

METHOD REGISTEREVENT
END_METHOD

METHOD UNREGISTEREVENT
END_METHOD

METHOD RESETHOMEPOS
END_METHOD

METHOD RESETHOMEPOS2
VAR_INPUT
	ERESETINFO : L_IE1P_Error;
END_VAR
END_METHOD

METHOD RESETHOMEPOSLOADENCODER
VAR_INPUT
	ERESETINFO : L_IE1P_Error;
END_VAR
END_METHOD

METHOD SETHOMEPOSDEPENDONMODESTATEINDEPENDENT : BOOL
VAR_INPUT
	EHOMEMODE : L_MC1P_HomeMode;
	LRPOSITION : LREAL;
	LROFFSETPOSITION : LREAL;
	EHOMEPOSINFO : L_IE1P_Error;
END_VAR
VAR_OUTPUT
	XERROR : BOOL;
	EERRORID : L_IE1P_Error;
END_VAR
END_METHOD

METHOD SETHOMEPOSITION
VAR_INPUT
	POSITION : LREAL;
	RELATIVE : BOOL;
	XRESTARTPOSITIONING : BOOL := FALSE;
END_VAR
END_METHOD

METHOD SETHOMEPOSITION2
VAR_INPUT
	POSITION : LREAL;
	RELATIVE : BOOL;
	XRESTARTPOSITIONING : BOOL := FALSE;
	EHOMEPOSINFO : L_IE1P_Error;
END_VAR
END_METHOD

METHOD SETHOMEPOSITIONWITHMODROUNDS
VAR_INPUT
	POSITION : LREAL;
	RELATIVE : BOOL;
	ROUNDS : LREAL;
	XRESTARTPOSITIONING : BOOL;
	EHOMEPOSINFO : L_IE1P_Error;
END_VAR
END_METHOD

METHOD ITFCHECKERRORRESETOCCURED : BOOL
VAR_IN_OUT
	RESETTIME : SYSTIME;
END_VAR
END_METHOD

METHOD ITFCLEARERROR : DWORD
VAR_INPUT
	ESEVERITY : L_IE1P_SeverityLevel;
	WERRORID : WORD;
	WCOMPID : WORD;
	DWINSTANCEID : DWORD := 0;
END_VAR
END_METHOD

METHOD ITFCLEARREACTION
VAR_INPUT
	EREACTION : L_IE1P_Reaction;
	DICLEARCOUNT : DINT;
	DWINSTANCEID : DWORD;
END_VAR
END_METHOD

METHOD ITFGETACTUALERRORCODE : DWORD
VAR_OUTPUT
	ESEVERITY : WORD;
END_VAR
END_METHOD

METHOD ITFREGISTERERRORINSTANCE : DWORD
END_METHOD

METHOD ITFRESETACTIVE : BOOL
END_METHOD

METHOD ITFRESETERROR : DWORD
VAR_INPUT
	ERRORHANDLE : SysTypes.RTS_IEC_HANDLE := 0;
END_VAR
END_METHOD

METHOD ITFRESETERRORREACTION
VAR_INPUT
	DWINSTANCEID : DWORD := 0;
END_VAR
END_METHOD

METHOD ITFSETERROR : DWORD
VAR_INPUT
	ESEVERITY : L_IE1P_SeverityLevel;
	WERRORID : WORD;
	WCOMPID : WORD;
	DWINSTANCEID : DWORD := 0;
	EREACTION : L_IE1P_Reaction;
END_VAR
END_METHOD

METHOD GETDIRECTION : WORD
VAR_INPUT
	VALUESOURCE : MC_SOURCE;
END_VAR
END_METHOD

METHOD GETMASTERERROR : BOOL
VAR_OUTPUT
	EERRORID : L_IE1P_Error;
END_VAR
END_METHOD

METHOD GETSTEADYSTATE : POINTER TO L_MC1P_SteadyState
END_METHOD

METHOD GETAXISFROMPOOL : POINTER TO AXIS_REF
VAR_INPUT
	WINDEX : WORD;
END_VAR
END_METHOD

METHOD CHECKINPOSITION
END_METHOD

METHOD SETINPOSITION
VAR_INPUT
	XDONE : BOOL;
	LRINTARGETPOSITION : LREAL;
END_VAR
END_METHOD

METHOD ACTIVATESS1
END_METHOD

METHOD CALCULATE_DECELERATION : LREAL
VAR_INPUT
	LRJERK : LREAL;
	LRTOTALTIME : LREAL;
	LRACTVEL : LREAL;
	LRTARGETVEL : LREAL;
	LRACCMAX : LREAL;
END_VAR
END_METHOD

METHOD CHECKLIMITERREQUESTS
END_METHOD

METHOD CHECKSLSCHANGES : BOOL
VAR_OUTPUT
	XLIMITERCONTROLCHANGED : BOOL;
	XSLSPARAMETERCHANGED : BOOL;
	XSLSNEWACTIVEDECELERATION : BOOL;
END_VAR
END_METHOD

METHOD CHECKSAFETYOPTIONAVAILABLE : BOOL
VAR_INPUT
	DWPRODUCTCODE : DWORD;
END_VAR
END_METHOD

METHOD LIMITSPEEDCONTROLLER
END_METHOD

METHOD PROCESSSSX
VAR_INPUT
	DWCONTROL : DWORD;
END_VAR
END_METHOD

METHOD UPDATEACTIVESLSSETVEL
VAR_INPUT
	LRVEL : LREAL;
END_VAR
END_METHOD

METHOD CHECKHWLIMITS : BOOL
END_METHOD

METHOD CHECKLIMITCHANGES : BOOL
VAR_OUTPUT
	XPOSSWLIMITCHANGED : BOOL;
	XNEGSWLIMITCHANGED : BOOL;
END_VAR
END_METHOD

METHOD CHECKMAXVALUES : BOOL
VAR_INPUT
	VELOCITY : LREAL;
	ACCELERATION : LREAL;
	JERK : LREAL;
END_VAR
END_METHOD

METHOD CHECKSWLIMITS : BOOL
VAR_INPUT
	XSETERRORSTOP : BOOL;
END_VAR
END_METHOD

METHOD DISABLESWLIMIT
VAR_INPUT
	XDISABLE : BOOL;
END_VAR
END_METHOD

METHOD GETACTDIRECTION : MC_DIRECTION
VAR_INPUT
	XCALCULATE : BOOL;
END_VAR
END_METHOD

METHOD GETSWLIMITSACTIVE : BOOL
END_METHOD

METHOD CALCCYCLELENGTH
END_METHOD

METHOD CALCULATESCALING : BOOL
END_METHOD

METHOD GETVIRTUAL : BOOL
END_METHOD

METHOD MACHINEDATACHANGED : BOOL
END_METHOD

METHOD WRITENEWMACHINEDATA
VAR_INPUT
	LRFEEDCONSTANTNEW : LREAL := 360.0;
	DWGEARDENOMINATORNEW : DWORD := 1;
	DWGEARNUMERATORNEW : DWORD := 1;
	DWADDGEARDENOMINATORNEW : DWORD := 1;
	DWADDGEARNUMERATORNEW : DWORD := 1;
	DWPOSRESOLUTIONNEW : DWORD := 65536;
	XORIENTATIONNEW : BOOL := FALSE;
	ETRAVERSINGRANGENEW : L_MC1P_TraversingRange := L_MC1P_TraversingRange.Limited;
	LRCYCLELENGTHNEW : LREAL := 360.0;
END_VAR
END_METHOD

METHOD COMPAREAXISNAME : BOOL
VAR_IN_OUT
	SAXISNAME : STRING;
END_VAR
END_METHOD

METHOD GETAXIS : POINTER TO AXIS_REF
END_METHOD

METHOD CALCSCALEFUNCTIONS
VAR_INPUT
	OFFSET : DWORD;
	INDEX : WORD;
END_VAR
END_METHOD

METHOD SETMACHINEDATAPARAMETER
END_METHOD

METHOD CALLCOMPFUNCTIONS
VAR_OUTPUT
	XCOMPERROR : BOOL;
END_VAR
END_METHOD

METHOD CALLFILTERFUNCTIONS
VAR_OUTPUT
	XFILTERERROR : BOOL;
END_VAR
END_METHOD

METHOD CHECKSETVALUESAVAILABLE
END_METHOD

METHOD RESETSETVALUESAVAILABLE
END_METHOD

METHOD RESTORESETVALUES
END_METHOD

METHOD SETCOMPITF : WORD
VAR_INPUT
	EINDEX : WORD;
	ITFCOMP : L_MC1P_ICompensationInterface;
END_VAR
END_METHOD

METHOD SETFILTERITF : WORD
VAR_INPUT
	EINDEX : WORD;
	ITFFILTER : L_MC1P_ISetvalueManipulationInterface;
	XFILTERINTERNALSET : BOOL;
END_VAR
END_METHOD

METHOD SETSETVALUESAVAILABLE
END_METHOD

METHOD SUSPENDSETVALUEFILTERCALL
VAR_INPUT
	XSUSPENDSETVALUEFILTERCALL : BOOL;
END_VAR
END_METHOD

METHOD ABORTACTIVEFUNCTION
END_METHOD

METHOD DRIVEQSP
END_METHOD

METHOD ERRORSTOP
END_METHOD

METHOD INTERNALSTOP : BOOL
VAR_INPUT
	XSTOP : BOOL;
	ESETSTATE : L_MC1P_AXIS_STATE;
	XPOSMODE : BOOL := FALSE;
	LRTARGETPOS : LREAL := 0;
	XABORTACTIVEFUNCTION : BOOL := TRUE;
END_VAR
VAR_IN_OUT
	XSTOPACTIVE : BOOL;
	XSTOPDONE : BOOL;
END_VAR
END_METHOD

METHOD MOVEBACKTOLASTSETPOS : BOOL
VAR_INPUT
	XSTOP : BOOL;
END_VAR
VAR_IN_OUT
	XSTOPACTIVE : BOOL;
	XSTOPDONE : BOOL;
END_VAR
END_METHOD

METHOD RAMPDOWN
END_METHOD

METHOD RAMPQSP
VAR_INPUT
	CALLEDFROMAPP : BOOL;
END_VAR
END_METHOD

METHOD RESETRAMPDOWN
END_METHOD

METHOD SETAXISSTOPINT : BOOL
VAR_INPUT
	XSTOP : BOOL;
	SCSTOPCMD : L_MC1P_StopOperation;
END_VAR
END_METHOD

METHOD SETFASTSTOPINT : BOOL
VAR_INPUT
	XSTOP : BOOL;
END_VAR
END_METHOD

METHOD SETSTANDSTILLSTATE
VAR_INPUT
	XRAMPDOWN : BOOL;
END_VAR
END_METHOD

METHOD STARTRAMPDOWN
END_METHOD

METHOD HLP_GETPARAMETER : BOOL
END_METHOD

METHOD HLP_GETPARAMETERPROPERTIES : BOOL
VAR_INPUT
	DIPARAMETER : DINT;
END_VAR
VAR_OUTPUT
	PPARAMADDR : POINTER TO BYTE := 0;
	EORDINALTYPE : L_MC1P_OrdinalType := L_MC1P_OrdinalType.otNONE;
	XREADWRITE : BOOL := FALSE;
	LRUNITFACTOR : LREAL := 1.0;
	LRDEFAULTVALUE : LREAL := 0.0;
	WVALUERANGES : WORD := 0;
	PVALUERANGES : POINTER TO L_MC1P_MinMaxValue := 0;
END_VAR
END_METHOD

METHOD HLP_INITPARREF
END_METHOD

METHOD HLP_READBOOLPARAMETER : BOOL
VAR_INPUT
	PARAMETER : DINT;
	PXVALUE : POINTER TO BOOL;
END_VAR
END_METHOD

METHOD HLP_READPARAMETER : BOOL
VAR_INPUT
	PARAMETER : DINT;
	PLRVALUE : POINTER TO LREAL;
END_VAR
END_METHOD

METHOD HLP_WRITEBOOLPARAMETER : BOOL
VAR_INPUT
	PARAMETER : DINT;
	PXVALUE : POINTER TO BOOL;
END_VAR
VAR_OUTPUT
	WERRORID : WORD;
END_VAR
END_METHOD

METHOD HLP_WRITEPARAMETER : BOOL
VAR_INPUT
	PARAMETER : DINT;
	PLRVALUE : POINTER TO LREAL;
END_VAR
VAR_OUTPUT
	WERRORID : WORD;
END_VAR
END_METHOD

METHOD AFTERREADINPUTS : INT
END_METHOD

METHOD AFTERWRITEOUTPUTS : INT
END_METHOD

METHOD BEFOREREADINPUTS : INT
END_METHOD

METHOD BEFOREWRITEOUTPUTS : INT
END_METHOD

METHOD CALCAFTERREADINPUTS : INT
END_METHOD

METHOD CALCAFTERWRITEOUTPUTS : INT
END_METHOD

METHOD CALCBEFOREREADINPUTS : INT
END_METHOD

METHOD CALCBEFOREWRITEOUTPUTS : INT
END_METHOD

METHOD FB_EXIT : BOOL
VAR_INPUT
	BINCOPYCODE : BOOL;
END_VAR
END_METHOD

METHOD INITFORSIMULATIONMODE : BOOL
VAR_INPUT
	WMODULETYPE : UINT;
	DWINSTANCE : UDINT;
	PCONNECTOR : POINTER TO IoConfigConnector;
END_VAR
END_METHOD

METHOD INITIALIZE : UDINT
VAR_INPUT
	WMODULETYPE : UINT;
	DWINSTANCE : UDINT;
	PCONNECTOR : POINTER TO IoConfigConnector;
END_VAR
END_METHOD

METHOD IODRVREADPARAMETER : UDINT
VAR_INPUT
	PCONNECTOR : POINTER TO IoConfigConnector;
	PPARAMETER : POINTER TO IoConfigParameter;
	PDATA : POINTER TO BYTE;
	DWBITSIZE : DWORD;
	DWBITOFFSET : DWORD;
END_VAR
END_METHOD

METHOD IODRVUPDATECONFIGURATION : UDINT
VAR_INPUT
	PCONNECTORLIST : POINTER TO IoConfigConnector;
	NCOUNT : DINT;
END_VAR
END_METHOD

METHOD IODRVUPDATEMAPPING : UDINT
VAR_INPUT
	PTASKMAPLIST : POINTER TO IoConfigTaskMap;
	NCOUNT : DINT;
END_VAR
END_METHOD

METHOD IODRVWRITEPARAMETER : UDINT
VAR_INPUT
	PCONNECTOR : POINTER TO IoConfigConnector;
	PPARAMETER : POINTER TO IoConfigParameter;
	PDATA : POINTER TO BYTE;
	DWBITSIZE : DWORD;
	DWBITOFFSET : DWORD;
END_VAR
END_METHOD

METHOD FB_INIT : BOOL
VAR_INPUT
	BINITRETAINS : BOOL;
	BINCOPYCODE : BOOL;
END_VAR
END_METHOD

METHOD FUNCTIONSUPPORTEDBYAXIS : BOOL
VAR_INPUT
	FUNID : L_MC1P_AxisFunction;
	XORIGINDEVICE : BOOL;
END_VAR
END_METHOD

METHOD GETDELAYFORFASTOUTPUTCALCULATION : LREAL
VAR_INPUT
	EVALUESOURCE : MC_SOURCE;
END_VAR
END_METHOD

METHOD GETINDEXOFENCODERCRC : WORD
END_METHOD

METHOD GETINDEXOFERRORCODE : DINT
END_METHOD

METHOD GETINDEXOFPOSCTRLADAPTVALUE
VAR_INPUT
	WSELECTION : WORD;
END_VAR
VAR_OUTPUT
	WINDEX : WORD;
	BYSUBINDEX : BYTE;
	BYSIZE : BYTE;
END_VAR
END_METHOD

METHOD GETINDEXOFSPEEDCTRLADAPTVALUE
VAR_INPUT
	WSELECTION : WORD;
END_VAR
VAR_OUTPUT
	WINDEX : WORD;
	BYSUBINDEX : BYTE;
	BYSIZE : BYTE;
END_VAR
END_METHOD

METHOD GETMAGNETISATIONFINISHED : BOOL
END_METHOD

METHOD GETMAXTORQUE : LREAL
END_METHOD

METHOD GETREFERENCETORQUE : LREAL
END_METHOD

METHOD GETTPDELAYFORFASTINPUTCALCULATION : LREAL
END_METHOD

METHOD GETVPPMAXVALUE : LREAL
END_METHOD

METHOD SETSPEEDCTRLLIMITATION : BOOL
VAR_INPUT
	XLIMIT : BOOL;
END_VAR
END_METHOD

METHOD SUPPORTLIMITSPEEDCONTROLLER : BOOL
VAR_OUTPUT
	WINDEX : WORD;
	BYSUBINDEX : BYTE;
	BYSIZE : BYTE;
END_VAR
END_METHOD

METHOD SUPPORTMFE : BOOL
END_METHOD

METHOD CALCDISTANCE : LREAL
VAR_INPUT
	LRROUNDSACT : LREAL;
	LRROUNDSSET : LREAL;
	LRPOSACT : LREAL;
	LRPOSSET : LREAL;
END_VAR
VAR_IN_OUT
	AXIS : AXIS_REF;
END_VAR
END_METHOD

METHOD CALCTARGETPOS : LREAL
VAR_INPUT
	LRROUNDSACT : LREAL;
	LRROUNDSSET : LREAL;
	LRPOSACT : LREAL;
	LRPOSSET : LREAL;
END_VAR
VAR_OUTPUT
	EDIR : MC_DIRECTION;
END_VAR
VAR_IN_OUT
	AXIS : AXIS_REF;
END_VAR
END_METHOD

METHOD SETPOSRECOVERYDATA
VAR_INPUT
	XACTIVATE : BOOL;
	LRVEL : LREAL;
	LRACC : LREAL;
	LRDEC : LREAL;
	LRJERK : LREAL;
END_VAR
END_METHOD

(* ---- AXIS_REF_9400HL.fb ---- *)
FUNCTION_BLOCK AXIS_REF_9400HL EXTENDS _AXIS_REF_9400HL
VAR
	PARA_AXIS_REF_9400HL : L_MC1P_ParaInterface_AXIS_REF_9400HL;
END_VAR
END_FUNCTION_BLOCK

METHOD FB_INIT : BOOL
VAR_INPUT
	BINITRETAINS : BOOL;
	BINCOPYCODE : BOOL;
END_VAR
END_METHOD

(* ---- AXIS_REF_9400HL_CAN.fb ---- *)
FUNCTION_BLOCK AXIS_REF_9400HL_CAN EXTENDS _AXIS_REF_9400HL_CAN
VAR
	PARA_AXIS_REF_9400HL_CAN : L_MC1P_ParaInterface_AXIS_REF_9400HL_CAN;
END_VAR
END_FUNCTION_BLOCK

METHOD FB_INIT : BOOL
VAR_INPUT
	BINITRETAINS : BOOL;
	BINCOPYCODE : BOOL;
END_VAR
END_METHOD

(* ---- AXIS_REF_ENC_BPB.fb ---- *)
FUNCTION_BLOCK AXIS_REF_ENC_BPB EXTENDS _AXIS_REF_ENC_BPB
VAR
	PARA_AXIS_REF_ENC_BPB : L_MC1P_ParaInterface_AXIS_REF_ENC_BPB;
END_VAR
END_FUNCTION_BLOCK

METHOD FB_INIT : BOOL
VAR_INPUT
	BINITRETAINS : BOOL;
	BINCOPYCODE : BOOL;
END_VAR
END_METHOD

(* ---- AXIS_REF_ENC_FREE.fb ---- *)
FUNCTION_BLOCK AXIS_REF_ENC_FREE EXTENDS _AXIS_REF_ENC_FREE
VAR
	PARA_AXIS_REF_ENC_FREE : L_MC1P_ParaInterface_AXIS_REF_ENC_FREE;
END_VAR
END_FUNCTION_BLOCK

METHOD FB_INIT : BOOL
VAR_INPUT
	BINITRETAINS : BOOL;
	BINCOPYCODE : BOOL;
END_VAR
END_METHOD

(* ---- AXIS_REF_ENC_I500_ECAT.fb ---- *)
FUNCTION_BLOCK AXIS_REF_ENC_I500_ECAT EXTENDS _AXIS_REF_ENC_i500_ECAT
VAR
	PARA_AXIS_REF_ENC_I500_ECAT : L_MC1P_ParaInterface_AXIS_REF_ENC_i500_ECAT;
END_VAR
END_FUNCTION_BLOCK

METHOD FB_INIT : BOOL
VAR_INPUT
	BINITRETAINS : BOOL;
	BINCOPYCODE : BOOL;
END_VAR
END_METHOD

(* ---- AXIS_REF_ENC_I900_DRIVE.fb ---- *)
FUNCTION_BLOCK AXIS_REF_ENC_I900_DRIVE EXTENDS _AXIS_REF_ENC_i900_Target
VAR
	PARA_AXIS_REF_ENC_I900_DRIVE : L_MC1P_ParaInterface_AXIS_REF_ENC_i900_DRIVE;
END_VAR
END_FUNCTION_BLOCK

METHOD FB_INIT : BOOL
VAR_INPUT
	BINITRETAINS : BOOL;
	BINCOPYCODE : BOOL;
END_VAR
END_METHOD

(* ---- AXIS_REF_ENC_I900_DRIVE_CIA.fb ---- *)
FUNCTION_BLOCK AXIS_REF_ENC_I900_DRIVE_CIA EXTENDS _AXIS_REF_ENC_i900_CiA
VAR
	PARA_AXIS_REF_ENC_I900_DRIVE_CIA : L_MC1P_ParaInterface_AXIS_REF_ENC_i900_DRIVE_CIA;
END_VAR
END_FUNCTION_BLOCK

METHOD FB_INIT : BOOL
VAR_INPUT
	BINITRETAINS : BOOL;
	BINCOPYCODE : BOOL;
END_VAR
END_METHOD

(* ---- AXIS_REF_ENC_I900_ECAT.fb ---- *)
FUNCTION_BLOCK AXIS_REF_ENC_I900_ECAT EXTENDS _AXIS_REF_ENC_i900_ECAT
VAR
	PARA_AXIS_REF_ENC_I900_ECAT : L_MC1P_ParaInterface_AXIS_REF_ENC_i900_ECAT;
END_VAR
END_FUNCTION_BLOCK

METHOD FB_INIT : BOOL
VAR_INPUT
	BINITRETAINS : BOOL;
	BINCOPYCODE : BOOL;
END_VAR
END_METHOD

(* ---- AXIS_REF_ENC_IO_ETC.fb ---- *)
FUNCTION_BLOCK AXIS_REF_ENC_IO_ETC EXTENDS _AXIS_REF_ENC_IO_ETC
VAR
	PARA_AXIS_REF_ENC_IO_ETC : L_MC1P_ParaInterface_AXIS_REF_ENC_IO_ETC;
END_VAR
END_FUNCTION_BLOCK

METHOD FB_INIT : BOOL
VAR_INPUT
	BINITRETAINS : BOOL;
	BINCOPYCODE : BOOL;
END_VAR
END_METHOD

(* ---- AXIS_REF_ENC_UNIVERSAL.fb ---- *)
FUNCTION_BLOCK AXIS_REF_ENC_UNIVERSAL EXTENDS _AXIS_REF_Enc_Universal
VAR
	PARA_AXIS_REF_ENC_UNIVERSAL : L_MC1P_ParaInterface_AXIS_REF_ENC_UNIVERSAL;
END_VAR
END_FUNCTION_BLOCK

METHOD FB_INIT : BOOL
VAR_INPUT
	BINITRETAINS : BOOL;
	BINCOPYCODE : BOOL;
END_VAR
END_METHOD

(* ---- AXIS_REF_GENERIC.fb ---- *)
FUNCTION_BLOCK AXIS_REF_GENERIC EXTENDS _AXIS_REF_GENERIC
VAR
	PARA_AXIS_REF_GENERIC : L_MC1P_ParaInterface_AXIS_REF_GENERIC;
END_VAR
END_FUNCTION_BLOCK

METHOD FB_INIT : BOOL
VAR_INPUT
	BINITRETAINS : BOOL;
	BINCOPYCODE : BOOL;
END_VAR
END_METHOD

(* ---- AXIS_REF_I500_CAN.fb ---- *)
FUNCTION_BLOCK AXIS_REF_I500_CAN EXTENDS _AXIS_REF_i500_CAN
VAR
	PARA_AXIS_REF_I500_CAN : L_MC1P_ParaInterface_AXIS_REF_i500_CAN;
END_VAR
END_FUNCTION_BLOCK

METHOD FB_INIT : BOOL
VAR_INPUT
	BINITRETAINS : BOOL;
	BINCOPYCODE : BOOL;
END_VAR
END_METHOD

(* ---- AXIS_REF_I500_ETC.fb ---- *)
FUNCTION_BLOCK AXIS_REF_I500_ETC EXTENDS _AXIS_REF_i500_ETC
VAR
	PARA_AXIS_REF_I500_ETC : L_MC1P_ParaInterface_AXIS_REF_i500_ETC;
END_VAR
END_FUNCTION_BLOCK

METHOD FB_INIT : BOOL
VAR_INPUT
	BINITRETAINS : BOOL;
	BINCOPYCODE : BOOL;
END_VAR
END_METHOD

(* ---- AXIS_REF_I700.fb ---- *)
FUNCTION_BLOCK AXIS_REF_I700 EXTENDS _AXIS_REF_i700
VAR
	PARA_AXIS_REF_I700 : L_MC1P_ParaInterface_AXIS_REF_i700;
END_VAR
END_FUNCTION_BLOCK

METHOD FB_INIT : BOOL
VAR_INPUT
	BINITRETAINS : BOOL;
	BINCOPYCODE : BOOL;
END_VAR
END_METHOD

(* ---- AXIS_REF_I700_SLOT1.fb ---- *)
FUNCTION_BLOCK AXIS_REF_I700_SLOT1 EXTENDS _AXIS_REF_i700_SLOT1
VAR
	PARA_AXIS_REF_I700_SLOT1 : L_MC1P_ParaInterface_AXIS_REF_i700_SLOT1;
END_VAR
END_FUNCTION_BLOCK

METHOD FB_INIT : BOOL
VAR_INPUT
	BINITRETAINS : BOOL;
	BINCOPYCODE : BOOL;
END_VAR
END_METHOD

(* ---- AXIS_REF_I750.fb ---- *)
FUNCTION_BLOCK AXIS_REF_I750 EXTENDS _AXIS_REF_i750
VAR
	PARA_AXIS_REF_I750 : L_MC1P_ParaInterface_AXIS_REF_i750;
END_VAR
END_FUNCTION_BLOCK

METHOD FB_INIT : BOOL
VAR_INPUT
	BINITRETAINS : BOOL;
	BINCOPYCODE : BOOL;
END_VAR
END_METHOD

(* ---- AXIS_REF_I900.fb ---- *)
FUNCTION_BLOCK AXIS_REF_I900 EXTENDS _AXIS_REF_i900
VAR
	PARA_AXIS_REF_I900 : L_MC1P_ParaInterface_AXIS_REF_i900;
END_VAR
END_FUNCTION_BLOCK

METHOD FB_INIT : BOOL
VAR_INPUT
	BINITRETAINS : BOOL;
	BINCOPYCODE : BOOL;
END_VAR
END_METHOD

(* ---- AXIS_REF_I900_CIAADV.fb ---- *)
FUNCTION_BLOCK AXIS_REF_I900_CIAADV EXTENDS _AXIS_REF_i900_CiaAdv
VAR
	PARA_AXIS_REF_I900_CIAADV : L_MC1P_ParaInterface_AXIS_REF_i900_CiaAdv;
END_VAR
END_FUNCTION_BLOCK

METHOD FB_INIT : BOOL
VAR_INPUT
	BINITRETAINS : BOOL;
	BINCOPYCODE : BOOL;
END_VAR
END_METHOD

(* ---- AXIS_REF_I900_DRIVE.fb ---- *)
FUNCTION_BLOCK AXIS_REF_I900_DRIVE EXTENDS _AXIS_REF_i900_Drive_Target
VAR
	PARA_AXIS_REF_I900_DRIVE : L_MC1P_ParaInterface_AXIS_REF_i900_DRIVE;
END_VAR
END_FUNCTION_BLOCK

METHOD FB_INIT : BOOL
VAR_INPUT
	BINITRETAINS : BOOL;
	BINCOPYCODE : BOOL;
END_VAR
END_METHOD

(* ---- AXIS_REF_I900_DRIVE_CIA.fb ---- *)
FUNCTION_BLOCK AXIS_REF_I900_DRIVE_CIA EXTENDS _AXIS_REF_i900_Drive_CiA
VAR
	PARA_AXIS_REF_I900_DRIVE_CIA : L_MC1P_ParaInterface_AXIS_REF_i900_DRIVE_CIA;
END_VAR
END_FUNCTION_BLOCK

METHOD FB_INIT : BOOL
VAR_INPUT
	BINITRETAINS : BOOL;
	BINCOPYCODE : BOOL;
END_VAR
END_METHOD

(* ---- AXIS_REF_UNIVERSAL.fb ---- *)
FUNCTION_BLOCK AXIS_REF_UNIVERSAL EXTENDS _AXIS_REF_Universal
VAR
	PARA_AXIS_REF_UNIVERSAL : L_MC1P_ParaInterface_AXIS_REF_UNIVERSAL;
END_VAR
END_FUNCTION_BLOCK

METHOD FB_INIT : BOOL
VAR_INPUT
	BINITRETAINS : BOOL;
	BINCOPYCODE : BOOL;
END_VAR
END_METHOD

(* ---- AXIS_REF_VIRTUAL.fb ---- *)
FUNCTION_BLOCK AXIS_REF_VIRTUAL EXTENDS AXIS_REF
VAR
	PARA_AXIS_REF_VIRTUAL : L_MC1P_ParaInterface_AXIS_REF_VIRTUAL;
END_VAR
END_FUNCTION_BLOCK

METHOD FB_INIT : BOOL
VAR_INPUT
	BINITRETAINS : BOOL;
	BINCOPYCODE : BOOL;
END_VAR
END_METHOD

(* ---- AXIS_REF_VIRTUALM_I900.fb ---- *)
FUNCTION_BLOCK AXIS_REF_VIRTUALM_I900 EXTENDS AXIS_REF
VAR
	PARA_AXIS_REF_VIRTUALM_I900 : L_MC1P_ParaInterface_AXIS_REF_VIRTUALM_i900;
END_VAR
END_FUNCTION_BLOCK

METHOD FB_INIT : BOOL
VAR_INPUT
	BINITRETAINS : BOOL;
	BINCOPYCODE : BOOL;
END_VAR
END_METHOD

(* ---- AXIS_REF_VMA.fb ---- *)
FUNCTION_BLOCK AXIS_REF_VMA EXTENDS _AXIS_REF_VMA
VAR
	PARA_AXIS_REF_VMA : L_MC1P_ParaInterface_AXIS_REF_VMA;
END_VAR
END_FUNCTION_BLOCK

METHOD FB_INIT : BOOL
VAR_INPUT
	BINITRETAINS : BOOL;
	BINCOPYCODE : BOOL;
END_VAR
END_METHOD

(* ---- GLOBALTEXTLIST.fb ---- *)
FUNCTION_BLOCK GLOBALTEXTLIST
VAR
	M_TEXTLISTFILE : STRING(255);
	_STNAMESPACE : STRING;
END_VAR
END_FUNCTION_BLOCK

(* ---- IMAGEPOOL.fb ---- *)
FUNCTION_BLOCK IMAGEPOOL
VAR
	M_STNAMESPACE : STRING(80);
	M_STHELPVARID : STRING;
	M_STHELPVARPATH : STRING(255);
	M_STHELP : STRING;
	M_REGISTERIMAGES : BOOL := TRUE;
END_VAR
END_FUNCTION_BLOCK

METHOD FB_INIT : BOOL
VAR_INPUT
	BINITRETAINS : BOOL;
	BINCOPYCODE : BOOL;
END_VAR
END_METHOD

METHOD FB_REINIT : BOOL
END_METHOD

METHOD FB_EXIT : BOOL
VAR_INPUT
	BINCOPYCODE : BOOL;
END_VAR
END_METHOD

(* ---- L_MB1P_TPCONVERTTP.fb ---- *)
FUNCTION_BLOCK L_MB1P_TPCONVERTTP
VAR_INPUT
	XENABLE : BOOL;
	XTPRECEIVE : BOOL;
	LRACTTPPOSIN : LREAL;
	LRCYCPOSTPAXIS : LREAL;
	LRCYCPOSTARGETAXIS : LREAL;
	LRCYCLELENGTHTPAXIS : LREAL;
	LRCYCLELENGTHTARGETAXIS : LREAL;
END_VAR
VAR_OUTPUT
	XTPRECEIVED : BOOL;
	LRTPACTPOS : LREAL;
	XERROR : BOOL;
	EERRORID : L_IE1P_Error;
END_VAR
VAR
	LRPOSFIFOX : ARRAY [1..20] OF LREAL := [10(0)];
	LRPOSFIFOREG : ARRAY [1..20] OF LREAL := [10(0)];
	BYCOUNTER : INT := 1;
	LRSTACKDIFFERENCE : LREAL;
	LRTPDELTAINMS : LREAL;
	LRDELTAPCT : LREAL;
	XTPRECEIVEDOLD : BOOL;
	LRTEMP : LREAL;
	IDIRECTION : INT;
	LRACTTPPOSIN_OLD : LREAL;
	XWAIT : BOOL;
	XWAIT_OLD : BOOL;
	LRACTTPPOSIN_INT : LREAL;
	R_TRIG1 : R_TRIG;
END_VAR
END_FUNCTION_BLOCK

METHOD SEARCHINSTACKNEGATIVE
END_METHOD

METHOD SEARCHINSTACKPOSITIVE
END_METHOD

(* ---- L_MB1P_TPTIMESTAMPTOPOS.fb ---- *)
FUNCTION_BLOCK L_MB1P_TPTIMESTAMPTOPOS
VAR_INPUT
	XENABLE : BOOL;
	XTPRECEIVE : BOOL;
	DWTPTIMESTAMP : DWORD;
	LRACTPOSIN : LREAL;
	LRCYCLELENGTH : LREAL;
	DWDELAYACTPOS : DWORD;
END_VAR
VAR_OUTPUT
	XBUSY : BOOL;
	XERROR : BOOL;
	EERRORID : L_IE1P_Error;
	XTPRECEIVED : BOOL;
	LRTPACTPOS : LREAL;
END_VAR
VAR
	XENABLEOLD : BOOL;
	WACTIDX : WORD;
	ALRPOS : ARRAY [0..31] OF LREAL;
	DITIMESTAMPDIFF : DINT;
	DWACTDCTIME : DWORD;
	DWTASKYCLE_NS : DWORD;
	XINIT : BOOL := TRUE;
	LRBASE : LREAL;
	LRDIFF : LREAL;
	LRFACTOR : LREAL;
	LRCAPTURE : LREAL;
	UDIINTERVAL : UDINT;
	LRINTERVAL : LREAL;
	XTPRECEIVEOLD : BOOL;
	C_WMAXELEMENTS : WORD := 31;
END_VAR
END_FUNCTION_BLOCK

METHOD CALCTPPOS : LREAL
END_METHOD

(* ---- L_MC1P_ABORTTRIGGER_INTERNAL.fb ---- *)
FUNCTION_BLOCK L_MC1P_ABORTTRIGGER_INTERNAL EXTENDS L_MC1P_Template_IntFB
VAR_INPUT
	EXECUTE : BOOL;
	PAUSEACTIVETP : BOOL;
END_VAR
VAR_OUTPUT
	DONE : BOOL;
	BUSY : BOOL;
	ERROR : BOOL;
	ERRORID : L_IE1P_Error;
END_VAR
VAR
	PTPREF : POINTER TO L_MC1P_TPData;
	EXECUTEOLD : BOOL := FALSE;
	SNTPNUMBER : SINT;
END_VAR
END_FUNCTION_BLOCK

METHOD MAIN
VAR_IN_OUT
	AXIS : AXIS_REF;
	FBBASE : L_MC1P_Template_ForAxis;
	TRIGGERINPUT : MC_TRIGGER_REF;
END_VAR
END_METHOD

(* ---- L_MC1P_ADDOFFSETCYCLIC.fb ---- *)
FUNCTION_BLOCK L_MC1P_ADDOFFSETCYCLIC
VAR_INPUT
	LRSETPOS : LREAL;
	LRSETOFFSET : LREAL;
	ETRAVERSINGRANGE : L_MC1P_TraversingRange := L_MC1P_TraversingRange.Modulo;
	LRCYCLELENGTH : LREAL;
END_VAR
VAR_OUTPUT
	LRSETPOSOUT : LREAL;
	XERROR : BOOL;
	EERRORID : L_IE1P_Error;
END_VAR
VAR
	LRPOSDIFF : LREAL;
	LRPOS : LREAL;
	LRLENGTH : LREAL;
END_VAR
END_FUNCTION_BLOCK

(* ---- L_MC1P_AVERAGEFILTERSETVALUES.fb ---- *)
FUNCTION_BLOCK L_MC1P_AVERAGEFILTERSETVALUES EXTENDS L_MC1P_SetSetValueManipulator
VAR_INPUT
	WFILTERDEPTH : WORD;
	XMANIPULATETORQUE : BOOL := FALSE;
END_VAR
VAR_OUTPUT
	XINEQOUT : BOOL;
END_VAR
VAR
	WFILTERDEPTHINT : WORD := 20;
	CWFILTERDEPTHMAX : WORD := 1000;
	LRFILTERDEPTH : LREAL;
	LRINVFILTERDEPTH : LREAL;
	WCOUNTER : WORD;
	XERROR_CHECKINPUTDATA : BOOL;
	LRHOMINGOFFSETACT : LREAL;
	LRFILTEREDPOS : LREAL;
	AVERAGEFILTER : L_MC1P_TimeAverage;
	XMANIPULATETORQUEINT : BOOL := FALSE;
END_VAR
END_FUNCTION_BLOCK

METHOD CALCULATE2
VAR_IN_OUT
	AXIS : AXIS_REF;
END_VAR
END_METHOD

METHOD CALLCYCLIC2
VAR_IN_OUT
	AXIS : AXIS_REF;
END_VAR
END_METHOD

METHOD ENABLEINIT2
VAR_IN_OUT
	AXIS : Axis_REf;
END_VAR
END_METHOD

METHOD INITIALIZEFILTER
END_METHOD

METHOD LOADOFFSET2
VAR_INPUT
	OFFSET : LREAL;
END_VAR
VAR_IN_OUT
	AXIS : AXIS_REF;
END_VAR
END_METHOD

METHOD READINPUTS2
VAR_IN_OUT
	AXIS : AXIS_REF;
END_VAR
END_METHOD

(* ---- L_MC1P_AXIS_REF_POOL_2AXES.fb ---- *)
FUNCTION_BLOCK L_MC1P_AXIS_REF_POOL_2AXES
VAR_OUTPUT
	AXESPOOL : L_MC1P_IAXIS_REF_POOL;
END_VAR
VAR_IN_OUT
	AXIS1 : AXIS_REF;
	AXIS2 : AXIS_REF;
END_VAR
VAR
	AAXIS : ARRAY [1..2] OF POINTER TO AXIS_REF;
	WAXISCOUNT : WORD;
	AXISPOOLCOUNT : WORD;
END_VAR
END_FUNCTION_BLOCK

METHOD GETAXISFROMPOOL : POINTER TO AXIS_REF
VAR_INPUT
	WINDEX : WORD;
END_VAR
END_METHOD

(* ---- L_MC1P_AXIS_REF_POOL_3AXES.fb ---- *)
FUNCTION_BLOCK L_MC1P_AXIS_REF_POOL_3AXES
VAR_OUTPUT
	AXESPOOL : L_MC1P_IAXIS_REF_POOL;
END_VAR
VAR_IN_OUT
	AXIS1 : AXIS_REF;
	AXIS2 : AXIS_REF;
	AXIS3 : AXIS_REF;
END_VAR
VAR
	AAXIS : ARRAY [1..3] OF POINTER TO AXIS_REF;
	WAXISCOUNT : WORD;
	AXISPOOLCOUNT : WORD;
END_VAR
END_FUNCTION_BLOCK

METHOD GETAXISFROMPOOL : POINTER TO AXIS_REF
VAR_INPUT
	WINDEX : WORD;
END_VAR
END_METHOD

(* ---- L_MC1P_AXISBASICCONTROL.fb ---- *)
FUNCTION_BLOCK L_MC1P_AXISBASICCONTROL EXTENDS L_MC1P_Template_Licence_150
VAR_INPUT
	XENABLEINTERNALCONTROL : BOOL;
	XREGULATORON : BOOL;
	XRESETERROR : BOOL;
	XENABLEPOSITIVE : BOOL := TRUE;
	XENABLENEGATIVE : BOOL := TRUE;
	XDISABLESWLIMIT : BOOL := FALSE;
	LROVERRIDE : LREAL := 1.0;
	LROVERRIDEACC : LREAL := 1.0;
	LROVERRIDEJERK : LREAL := 1.0;
	XSTOP : BOOL;
	LRSTOPDEC : LREAL := 360000;
	LRSTOPJERK : LREAL := 0;
	XJOGGINGPOS : BOOL;
	XJOGGINGNEG : BOOL;
	LRJOGGINGSETVEL : LREAL := 3600;
	LRJOGGINGSETACC : LREAL := 36000;
	LRJOGGINGSETDEC : LREAL := 36000;
	LRJOGGINGSETJERK : LREAL := 0;
	XCONTINUOUSUPDATE : BOOL;
	XMOVEVELEXECUTE : BOOL;
	XMOVEABSEXECUTE : BOOL;
	XMOVERELEXECUTE : BOOL;
	XHALT : BOOL;
	LRSETPOS_DIST : LREAL;
	LRSETVEL : LREAL := 3600;
	LRSETACC : LREAL := 36000;
	LRSETDEC : LREAL := 36000;
	LRSETJERK : LREAL := 0;
	ESETDIRECTION : MC_DIRECTION := MC_DIRECTION.mcPositiveDirection;
	XHOMEEXECUTE : BOOL;
	LRHOMEPOSITION : LREAL;
	XUSEHOMEEXTPARAMETER : BOOL;
	SCHOMEEXTPARAMETER : L_MC1P_HomeParameter;
	SCHOMEEXTTP : MC_TRIGGER_REF;
	XHOMEABSSWITCH : BOOL;
END_VAR
VAR_OUTPUT
	XINTERNALCONTROLACTIVE : BOOL;
	XERROR : BOOL;
	EERRORID : L_IE1P_Error;
	XFUNBUSY : BOOL;
	XFUNDONE : BOOL;
	XFUNCOMMANDABORTED : BOOL;
	EFUNSTATEACT : L_MC1P_ABC_State;
	ECONTROLMODE : L_MC1P_ControlMode;
	XISHOMED : BOOL;
	XHWLIMITSWITCHNEG : BOOL;
	XHWLIMITSWITCHPOS : BOOL;
	XSWLIMITENABLED : BOOL;
	XSWLIMITSWITCHNEG : BOOL;
	XSWLIMITSWITCHPOS : BOOL;
	EAXISTYPE : L_MC1P_DriveType;
	EAXISSTATE : L_MC1P_AXIS_STATE := L_MC1P_AXIS_STATE.Disabled;
	XAXISREADY : BOOL;
	XAXISENABLED : BOOL;
	XAXISWARNING : BOOL;
	XAXISERROR : BOOL;
	EAXISERRORID : L_IE1P_Error;
	XDRIVEWARNING : BOOL;
	XDRIVEERROR : BOOL;
	DWDRIVEERRORID : DWORD;
	LRACTPOS : LREAL;
	LRACTVEL : LREAL;
	LRSETPOSOUT : LREAL;
	LRSETVELOUT : LREAL;
	LRACTFOLLOWINGERROR : LREAL;
	XCONSTANTVELOCITY : BOOL;
	XACCELERATING : BOOL;
	XDECELERATING : BOOL;
	XDIRECTIONPOSITIVE : BOOL;
	XDIRECTIONNEGATIVE : BOOL;
	XINPOSITION : BOOL;
	XAXISAVAILABLE : BOOL;
	XSTANDSTILLSETVELOCITY : BOOL;
	XSTANDSTILLACTVELOCITY : BOOL;
	XAXISREADYTOSWITCHON : BOOL;
	XAXISREADYFORMOTION : BOOL;
END_VAR
VAR
	XREGULATORON_INT : BOOL;
	XRESETERROR_INT : BOOL;
	XENABLEPOSITIVE_INT : BOOL;
	XENABLENEGATIVE_INT : BOOL;
	XDISABLESWLIMIT_INT : BOOL;
	LROVERRIDE_INT : LREAL := 1.0;
	LROVERRIDEACC_INT : LREAL := 1.0;
	LROVERRIDEJERK_INT : LREAL := 1.0;
	XSTOP_INT : BOOL;
	LRSTOPDEC_INT : LREAL;
	LRSTOPJERK_INT : LREAL;
	XHALT_INT : BOOL;
	XJOGGINGPOS_INT : BOOL;
	XJOGGINGNEG_INT : BOOL;
	LRJOGGINGSETVEL_INT : LREAL;
	LRJOGGINGSETACC_INT : LREAL;
	LRJOGGINGSETDEC_INT : LREAL;
	LRJOGGINGSETJERK_INT : LREAL := 0;
	LRJOGGINGSETJERKDEC_INT : LREAL := 0;
	LRJOGGINGSETJERKDECAPP : LREAL := 0;
	XMOVEVELEXECUTE_INT : BOOL;
	XMOVEABSEXECUTE_INT : BOOL;
	XMOVERELEXECUTE_INT : BOOL;
	XCONTINUOUSUPDATE_INT : BOOL;
	LRSETPOS_DIST_INT : LREAL;
	LRSETVEL_INT : LREAL;
	LRSETACC_INT : LREAL;
	LRSETDEC_INT : LREAL;
	LRSETJERK_INT : LREAL;
	LRSETJERKDEC_INT : LREAL := 0;
	LRSETJERKDECAPP : LREAL := 0;
	ESETDIRECTION_INT : MC_DIRECTION;
	XHOMEEXECUTE_INT : BOOL;
	LRHOMEPOSITION_INT : LREAL;
	XHOMEEXTERNALVALUES_INT : BOOL;
	SCHOMEEXTPARAMETER_INT : L_MC1P_HomeParameter;
	XDISABLEMOVEFUNEXEC : BOOL;
	XINTERNALCONTROLVISU : BOOL;
	XDISABLEMOVEFUN : BOOL;
	XDISABLEHOMEFUN : BOOL;
	XDISABLEPOWERFUN : BOOL;
	XDISABLEPOWERCALL : BOOL;
	XVISUMOVEFUN : BOOL;
	XVISUHOMEFUN : BOOL;
	XVISUPOWFUN : BOOL;
	ABC : REFERENCE TO L_MC1P_AxisBasicControl_Internal;
	DATA : L_MC1P_AxisBasicControlInstanceData;
	FBBASEOLD : POINTER TO L_MC1P_Template_ForAxis;
	_USEQSP : BOOL := FALSE;
	DISABLEHOMEFUN : BOOL;
	DISABLEMOVEFUN : BOOL;
	DISABLEMOVEFUNEXEC : BOOL;
	DISABLEPOWERCALL : BOOL;
	DISABLEPOWERFUN : BOOL;
	LRJOGGINGSETJERKDEC : LREAL;
	LRSETJERKDEC : LREAL;
	USEQSP : BOOL;
END_VAR
END_FUNCTION_BLOCK

(* ---- L_MC1P_AXISBASICCONTROL_INTERNAL.fb ---- *)
FUNCTION_BLOCK L_MC1P_AXISBASICCONTROL_INTERNAL EXTENDS L_MC1P_Template_IntFB
VAR_INPUT
	XDISABLEPOWERCALL : BOOL;
	XREGULATORON : BOOL;
	XRESETERROR : BOOL;
	XENABLEPOSITIVE : BOOL := TRUE;
	XENABLENEGATIVE : BOOL := TRUE;
	XDISABLESWLIMIT : BOOL;
	LROVERRIDE : LREAL := 1.0;
	LROVERRIDEACC : LREAL := 1.0;
	LROVERRIDEJERK : LREAL := 1.0;
	XSTOP : BOOL;
	LRSTOPDEC : LREAL;
	LRSTOPJERK : LREAL;
	XJOGGINGPOS : BOOL;
	XJOGGINGNEG : BOOL;
	LRJOGGINGSETVEL : LREAL := 3600;
	LRJOGGINGSETACC : LREAL := 36000;
	LRJOGGINGSETDEC : LREAL := 36000;
	LRJOGGINGSETJERK : LREAL := 0;
	LRJOGGINGSETJERKDEC : LREAL := 0;
	XCONTINUOUSUPDATE : BOOL;
	XFINISHPOSITIONING : BOOL;
	XQSPAPPLICATION : BOOL;
	XHALT : BOOL;
	XABORT : BOOL;
	XMOVEVELEXECUTE : BOOL;
	XMOVEABSEXECUTE : BOOL;
	XMOVERELEXECUTE : BOOL;
	LRSETPOS_DIST : LREAL;
	LRSETVEL : LREAL := 3600;
	LRSETACC : LREAL := 36000;
	LRSETDEC : LREAL := 36000;
	LRSETJERK : LREAL := 0;
	LRSETJERKDEC : LREAL := 0;
	ESETDIRECTION : MC_DIRECTION := MC_DIRECTION.mcPositiveDirection;
	XHOMEEXECUTE : BOOL;
	LRHOMEPOSITION : LREAL;
	XUSEHOMEEXTPARAMETER : BOOL;
	SCHOMEEXTPARAMETER : L_MC1P_HomeParameter;
	SCHOMEEXTTP : MC_TRIGGER_REF;
	XHOMEABSSWITCH : BOOL;
	XRESETHOMEPOSITION : BOOL;
	WCALLEDINCYCLE : WORD;
	XQSPDRIVEDONE : BOOL;
	XMOVEVELENABLEOFFSETVEL : BOOL;
	LRMOVEVELOFFSETVEL : LREAL;
	XUSEABORTBEHAVIOURFORTM : BOOL;
	LRABORTDEC : LREAL;
	LRABORTJERK : LREAL;
END_VAR
VAR_OUTPUT
	ECONTROLMODE : L_MC1P_ControlMode;
	XISHOMED : BOOL;
	XHWLIMITSWITCHNEG : BOOL;
	XHWLIMITSWITCHPOS : BOOL;
	XSWLIMITENABLED : BOOL;
	XSWLIMITSWITCHNEG : BOOL;
	XSWLIMITSWITCHPOS : BOOL;
	EAXISTYPE : L_MC1P_DriveType;
	EAXISSTATE : L_MC1P_AXIS_STATE := L_MC1P_AXIS_STATE.Disabled;
	XAXISREADY : BOOL;
	XAXISENABLED : BOOL;
	XAXISWARNING : BOOL;
	XAXISERROR : BOOL;
	EAXISERRORID : L_IE1P_Error;
	XDRIVEWARNING : BOOL;
	XDRIVEERROR : BOOL;
	DWDRIVEERRORID : DWORD;
	LRACTPOS : LREAL;
	LRACTVEL : LREAL;
	LRSETPOSOUT : LREAL;
	LRSETVELOUT : LREAL;
	LRACTFOLLOWINGERROR : LREAL;
	XCONSTANTVELOCITY : BOOL;
	XACCELERATING : BOOL;
	XDECELERATING : BOOL;
	XDIRECTIONPOSITIVE : BOOL;
	XDIRECTIONNEGATIVE : BOOL;
	XINPOSITION : BOOL;
	XAXISAVAILABLE : BOOL;
	XSTANDSTILLSETVELOCITY : BOOL;
	XSTANDSTILLACTVELOCITY : BOOL;
	XAXISREADYTOSWITCHON : BOOL;
	XAXISREADYFORMOTION : BOOL;
END_VAR
VAR
	ABCFUNID : WORD;
	FBSTOP : L_MC1P_Stop_Internal;
	FBHALT : L_MC1P_Halt_Internal;
	FBABORT : L_MC1P_Halt_Internal;
	FBHOME : L_MC1P_Home_Internal;
	FBJOG : L_MC1P_ManualJog_Internal;
	FBMOVEABS : L_MC1P_MoveAbsolute_Inernal;
	FBMOVEVEL : L_MC1P_MoveVelocity_Internal;
	FBMOVEREL : L_MC1P_MoveRelative_Internal;
	FBFINISHPOSITIONING : L_MC1P_FinishPositioning_internal;
	PBDUMMY : POINTER TO BOOL;
	XCONTROLLEDBYAXIS : BOOL;
	XCALLEDBYAXIS : BOOL;
	XUPDATESTATE : BOOL;
	XUPDATECONTROL : BOOL;
	XDISABLEMOVEFUNEXEC : BOOL;
	XDISABLEINTERNALCALLOFMOVEFUNCTIONS : BOOL;
	ETMPHOMEMODE : L_MC1P_HomeMode;
	LRTMPOFFSETPOSITION : LREAL;
	AXISCONTROL : BOOL;
	CALLEDBYAXIS : BOOL;
	DISABLEMOVEFUNEXEC : BOOL;
END_VAR
END_FUNCTION_BLOCK

METHOD BASEITFCHANGED
VAR_INPUT
	FBBASEOLD : POINTER TO POINTER TO L_MC1P_Template_ForAxis;
END_VAR
VAR_IN_OUT
	AXIS : AXIS_REF;
	FBBASE : L_MC1P_Template_ForAxis;
	DATA : L_MC1P_AxisBasicControlInstanceData;
END_VAR
END_METHOD

METHOD CALLMOVEFB : BOOL
VAR_IN_OUT
	AXIS : AXIS_REF;
	DATA : L_MC1P_AxisBasicControlInstanceData;
END_VAR
END_METHOD

METHOD EXITSTATE
VAR_IN_OUT
	AXIS : AXIS_REF;
	DATA : L_MC1P_AxisBasicControlInstanceData;
END_VAR
END_METHOD

METHOD MAIN
VAR_IN_OUT
	AXIS : AXIS_REF;
	FBBASE : L_MC1P_Template_ForAxis;
	DATA : L_MC1P_AxisBasicControlInstanceData;
END_VAR
END_METHOD

METHOD RESET
VAR_IN_OUT
	DATA : L_MC1P_AxisBasicControlInstanceData;
END_VAR
END_METHOD

METHOD RESETACTIVEINSTANCE : WORD
END_METHOD

METHOD SETACTIVEINSTANCE : WORD
END_METHOD

METHOD STATEMACHINE
VAR_IN_OUT
	AXIS : AXIS_REF;
	DATA : L_MC1P_AxisBasicControlInstanceData;
END_VAR
END_METHOD

(* ---- L_MC1P_AXISBASICCONTROLV2.fb ---- *)
FUNCTION_BLOCK L_MC1P_AXISBASICCONTROLV2 EXTENDS L_MC1P_Template_Licence_150
VAR_INPUT
	XENABLEINTERNALCONTROL : BOOL;
	XENABLEOPERATION : BOOL;
	XRESETERROR : BOOL;
	XENABLEPOSITIVE : BOOL := TRUE;
	XENABLENEGATIVE : BOOL := TRUE;
	XDISABLESWLIMIT : BOOL := FALSE;
	LROVERRIDE : LREAL := 1.0;
	LROVERRIDEACC : LREAL := 1.0;
	LROVERRIDEJERK : LREAL := 1.0;
	XQSPAPPLICATION : BOOL;
	XHALT : BOOL;
	XABORT : BOOL;
	XJOGPOS : BOOL;
	XJOGNEG : BOOL;
	XCONTINUOUSUPDATE : BOOL;
	XFINISHPOSITIONING : BOOL;
	XMOVEVELEXECUTE : BOOL;
	XMOVEABSEXECUTE : BOOL;
	XMOVERELEXECUTE : BOOL;
	LRPOS_DIST : LREAL := 0;
	LRVEL : LREAL := 3600;
	LRACC : LREAL := 36000;
	LRDEC : LREAL := 36000;
	LRJERK : LREAL := 0;
	EDIRECTION : MC_DIRECTION := MC_DIRECTION.mcPositiveDirection;
	XHOMEEXECUTE : BOOL;
	SCHOMEEXTTP : MC_TRIGGER_REF;
	XHOMEABSSWITCH : BOOL;
	XRESETHOMEPOSITION : BOOL;
END_VAR
VAR_OUTPUT
	XINTERNALCONTROLACTIVE : BOOL;
	XERROR : BOOL;
	EERRORID : L_IE1P_Error;
	XFUNBUSY : BOOL;
	XFUNDONE : BOOL;
	XFUNCOMMANDABORTED : BOOL;
	EFUNSTATEACT : L_MC1P_ABC_State := L_MC1P_ABC_State.Standby;
	ECONTROLMODE : L_MC1P_ControlMode := L_MC1P_ControlMode.PosCtrlDrive;
	XISHOMED : BOOL;
	XHWLIMITSWITCHNEG : BOOL;
	XHWLIMITSWITCHPOS : BOOL;
	XSWLIMITENABLED : BOOL;
	XSWLIMITSWITCHNEG : BOOL;
	XSWLIMITSWITCHPOS : BOOL;
	EAXISTYPE : L_MC1P_DriveType := L_MC1P_DriveType.Virtual;
	EAXISSTATE : L_MC1P_AXIS_STATE := L_MC1P_AXIS_STATE.Disabled;
	XSTOACTIVE : BOOL;
	XREADYFOROPERATION : BOOL;
	XOPERATIONENABLED : BOOL;
	XREADYFORMOTION : BOOL;
	XAXISWARNING : BOOL;
	XAXISERROR : BOOL;
	EAXISERRORID : L_IE1P_Error;
	XDRIVEWARNING : BOOL;
	XDRIVEERROR : BOOL;
	DWDRIVEERRORID : DWORD;
	LRACTPOS : LREAL;
	LRACTVEL : LREAL;
	LRSETPOSOUT : LREAL;
	LRSETVELOUT : LREAL;
	LRACTFOLLOWINGERROR : LREAL;
	XINPOSITION : BOOL;
	XSTANDSTILLSETVELOCITY : BOOL;
	XSTANDSTILLACTVELOCITY : BOOL;
	XCONSTANTVELOCITY : BOOL;
	XACCELERATING : BOOL;
	XDECELERATING : BOOL;
	XDIRECTIONPOSITIVE : BOOL;
	XDIRECTIONNEGATIVE : BOOL;
	XAXISAVAILABLE : BOOL;
END_VAR
VAR
	_ITFOWNER : L_UBUP.L_UBUP_IFBPool;
	_XWHANDLE : __XWORD;
	_XOCCUPIED : BOOL;
	XENABLEOPERATION_INT : BOOL;
	XRESETERROR_INT : BOOL;
	XENABLEPOSITIVE_INT : BOOL;
	XENABLENEGATIVE_INT : BOOL;
	XDISABLESWLIMIT_INT : BOOL;
	LROVERRIDE_INT : LREAL;
	LROVERRIDEACC_INT : LREAL;
	LROVERRIDEJERK_INT : LREAL;
	XQSPAPPLICATION_INT : BOOL;
	XHALT_INT : BOOL;
	XABORT_INT : BOOL;
	XJOGPOS_INT : BOOL;
	XJOGNEG_INT : BOOL;
	XCONTINUOUSUPDATE_INT : BOOL;
	XFINISHPOSITIONING_INT : BOOL;
	XMOVEVELEXECUTE_INT : BOOL;
	XMOVEABSEXECUTE_INT : BOOL;
	XMOVERELEXECUTE_INT : BOOL;
	LRPOS_DIST_INT : LREAL;
	LRVEL_INT : LREAL;
	LRACC_INT : LREAL;
	LRDEC_INT : LREAL;
	LRJERK_INT : LREAL;
	EDIRECTION_INT : MC_DIRECTION;
	XHOMEEXECUTE_INT : BOOL;
	XRESETHOMEPOSITION_INT : BOOL;
	LRSETJERKDEC_INT : LREAL;
	LRJOGGINGSETJERKDEC_INT : LREAL;
	LRSETJERKDECAPP : LREAL;
	LRJOGGINGSETJERKDECAPP : LREAL;
	XDISABLEMOVEFUNEXEC : BOOL;
	XDISABLEPOWERCALL : BOOL;
	XINTERNALCONTROLVISU : BOOL;
	XDISABLEMOVEFUN : BOOL;
	XDISABLEHOMEFUN : BOOL;
	XDISABLEPOWERFUN : BOOL;
	XVISUMOVEFUN : BOOL;
	XVISUHOMEFUN : BOOL;
	XVISUPOWFUN : BOOL;
	LRMOVEVELOFFSETVELAPP : LREAL;
	XMOVEVELENABLEOFFSETVELAPP : BOOL;
	LRABORTDECAPP : LREAL;
	LRABORTJERKAPP : LREAL;
	XUSEABORTBEHAVIOURFORTM : BOOL;
	ABC : REFERENCE TO L_MC1P_AxisBasicControl_Internal;
	DATA : L_MC1P_AxisBasicControlInstanceData;
	FBBASEOLD : POINTER TO L_MC1P_Template_ForAxis;
	_DWOBJID : DWORD;
	CLASSID : DINT;
	DISABLEHOMEFUN : BOOL;
	DISABLEMOVEFUN : BOOL;
	DISABLEMOVEFUNEXEC : BOOL;
	DISABLEPOWERCALL : BOOL;
	DISABLEPOWERFUN : BOOL;
	INSTANCEPTR : POINTER TO BYTE;
	LRABORTDEC : LREAL;
	LRABORTJERK : LREAL;
	LRJOGGINGSETJERKDEC : LREAL;
	LRMOVEVELOFFSETVEL : LREAL;
	LRSETJERKDEC : LREAL;
	OBJECTID : DWORD;
	OCCUPIED : BOOL;
	REMAININGTIMEOFPROFILE : LREAL;
	REMAININGTIMEOFPROFILEAVAILABLE : BOOL;
	XMOVEVELENABLEOFFSETVEL : BOOL;
	XSPECIALABORTBEHAVIOR : BOOL;
END_VAR
END_FUNCTION_BLOCK

METHOD RESETABORT
END_METHOD

METHOD RESETFINISHPOSITIONING
END_METHOD

METHOD RESETHALT
END_METHOD

METHOD RESETHOMEEXECUTE
END_METHOD

METHOD RESETMOVEABSEXECUTE
END_METHOD

METHOD RESETMOVERELEXECUTE
END_METHOD

METHOD RESETMOVEVELEXECUTE
END_METHOD

METHOD FREE : BOOL
END_METHOD

METHOD OCCUPY : BOOL
VAR_INPUT
	ITFOWNER : L_UBUP.L_UBUP_IFBPool;
	XWHANDLE : __XWORD;
END_VAR
END_METHOD

METHOD REQUESTINTERFACE : BOOL
VAR_INPUT
	ID : DINT;
	PITFUNKNOWN : POINTER TO L_UBUP_IUnknown;
END_VAR
END_METHOD

METHOD FB_INIT : BOOL
VAR_INPUT
	BINITRETAINS : BOOL;
	BINCOPYCODE : BOOL;
END_VAR
END_METHOD

(* ---- L_MC1P_AXISCOMMAND.fb ---- *)
FUNCTION_BLOCK L_MC1P_AXISCOMMAND
VAR_INPUT
	COMMANDIN : USINT;
END_VAR
VAR_OUTPUT
	XCOMMANDBUSY : BOOL;
END_VAR
VAR
	XABORT : BOOL;
	COMMAND : REFERENCE TO USINT;
	COMMANDOLD : USINT;
	FB_BASE : L_MC1P_Template_ForAxis;
	C_CMDREADY : USINT := 0;
	C_CMDSTART : USINT := 1;
	C_CMDINPROGRESS : USINT := 2;
	C_CMDCANCELLED : USINT := 3;
	C_CMDNOACCESS : USINT := 4;
	C_CMDNOACCESSDISABLED : USINT := 5;
	C_CMDABORT : USINT := 16;
	C_CMDWORKING20 : USINT := 20;
	C_CMDWORKING40 : USINT := 40;
	C_CMDWORKING60 : USINT := 60;
	C_CMDWORKING80 : USINT := 80;
	C_CMDWRONGBRAKEMODE : USINT := 101;
	C_CMDSTOACTIVE : USINT := 102;
	C_CMDINVALIDPARAMETERSETTINGS : USINT := 103;
	C_CMDSTARTOUTSIDEPOSLIMITS : USINT := 104;
	C_CMDPOSRANGENOTSUFFICIENT : USINT := 105;
	C_CMDHOMEPOSREQUIRED : USINT := 106;
	C_CMDINVALIDPOSITIONLIMITS : USINT := 107;
	C_CMDVIRTUALMODENOTSUPPORTED : USINT := 120;
	BUSY : BOOL;
END_VAR
END_FUNCTION_BLOCK

METHOD ABORTING
END_METHOD

METHOD CALCSTATUS
VAR_IN_OUT
	AXIS : _AXIS_REF_REAL;
END_VAR
END_METHOD

METHOD EXECUTE
END_METHOD

METHOD MAIN
END_METHOD

METHOD READINPUTS
END_METHOD

METHOD RESETCOMMANDERRORSTATE : BOOL
VAR_IN_OUT
	AXIS : _AXIS_REF_REAL;
END_VAR
END_METHOD

METHOD RESETSTATUSPARAMETER
END_METHOD

METHOD SETINCTANCEINFO
VAR_INPUT
	PSINSTANCENAME : POINTER TO STRING;
	ERRORITFID : DWORD;
END_VAR
END_METHOD

METHOD UPDATEAXISPOINTER
VAR_INPUT
	PAXIS : POINTER TO AXIS_REF;
END_VAR
END_METHOD

METHOD UPDATECOMMANDINTERFACE
VAR_IN_OUT
	CMD : USINT;
END_VAR
END_METHOD

METHOD FB_INIT : BOOL
VAR_INPUT
	BINITRETAINS : BOOL;
	BINCOPYCODE : BOOL;
END_VAR
END_METHOD

(* ---- L_MC1P_AXISCOMMAND_BRAKEGRINDIN.fb ---- *)
FUNCTION_BLOCK L_MC1P_AXISCOMMAND_BRAKEGRINDIN EXTENDS L_MC1P_AxisCommand
VAR_INPUT
	PAXIS : POINTER TO _AXIS_REF_REAL;
	EMODE : L_MC1P_GrindInMode := L_MC1P_GrindInMode.CwCcw;
	LRMOTORSPEED : LREAL := 60.0;
	LRRAMPTIME : LREAL := 1.0;
	LRONTIME : LREAL := 0.5;
	LROFFTIME : LREAL := 0.5;
	WCYCLES : WORD := 4;
	USICONTROL : USINT;
END_VAR
VAR
	FB_BRAKEGRINDIN : L_MC1P_BrakeGrindIn_internal;
	STATUS_100 : LREAL;
	LRSTATUS : LREAL;
	C_WSTATESUCCESSFUL : WORD := 10;
	C_WSTATEABORTEDERROR : WORD := 8;
	C_WSTATEABORTEDUSER : WORD := 9;
END_VAR
END_FUNCTION_BLOCK

METHOD ABORTING
END_METHOD

METHOD EXECUTE
END_METHOD

METHOD READINPUTS
END_METHOD

METHOD RESETSTATUSPARAMETER
END_METHOD

METHOD UPDATEAXISPOINTER
VAR_INPUT
	PAXIS : POINTER TO AXIS_REF;
END_VAR
END_METHOD

(* ---- L_MC1P_AXISCOMMAND_BRAKETEST.fb ---- *)
FUNCTION_BLOCK L_MC1P_AXISCOMMAND_BRAKETEST EXTENDS L_MC1P_AxisCommand
VAR_INPUT
	PAXIS : POINTER TO _AXIS_REF_REAL;
END_VAR
VAR
	FB_BRAKETEST : L_MC1P_BrakeTest_internal;
	ACTPOSTHRESHOLD : INT;
	STATUS_100 : LREAL;
	LRSTATUS : LREAL;
	LRTIME : LREAL;
	C_WSTATESUCCESSFUL : WORD := 10;
	C_WSTATEFAILED : WORD := 11;
	C_WSTATEABORTEDERROR : WORD := 8;
	C_WSTATEABORTEDUSER : WORD := 9;
END_VAR
END_FUNCTION_BLOCK

METHOD ABORTING
END_METHOD

METHOD EXECUTE
END_METHOD

METHOD READINPUTS
END_METHOD

METHOD RESETSTATUSPARAMETER
END_METHOD

METHOD UPDATEAXISPOINTER
VAR_INPUT
	PAXIS : POINTER TO AXIS_REF;
END_VAR
END_METHOD

(* ---- L_MC1P_AXISCONNECTIONVIEWER.fb ---- *)
FUNCTION_BLOCK L_MC1P_AXISCONNECTIONVIEWER EXTENDS L_IF1P_FunctionConnectionViewer
END_FUNCTION_BLOCK

METHOD BUILDUPCONNECTIONTABLE : BOOL
END_METHOD

METHOD FINDCONNECTIONSOURCE : POINTER TO BYTE
VAR_INPUT
	PSLAVECONNECTOR : POINTER TO IoConfigConnector;
	UITYPE : UINT;
	UISUBDEVICE : UINT;
END_VAR
END_METHOD

METHOD FINDFUNCTION : L_IF1P_IFunctionConnection
VAR_INPUT
	PFUNCTIONCONNECTOR : POINTER TO IoConfigConnector;
END_VAR
VAR_OUTPUT
	UITYPE : UINT;
END_VAR
END_METHOD

METHOD GETCONNECTEDSLAVE : BOOL
END_METHOD

METHOD INITIALIZE : UDINT
VAR_INPUT
	WMODULETYPE : UINT;
	DWINSTANCE : UDINT;
	PCONNECTOR : POINTER TO IoConfigConnector;
END_VAR
END_METHOD

METHOD IODRVREADPARAMETER : UDINT
VAR_INPUT
	PCONNECTOR : POINTER TO IoConfigConnector;
	PPARAMETER : POINTER TO IoConfigParameter;
	PDATA : POINTER TO BYTE;
	DWBITSIZE : DWORD;
	DWBITOFFSET : DWORD;
END_VAR
END_METHOD

METHOD IODRVUPDATECONFIGURATION : UDINT
VAR_INPUT
	PCONNECTORLIST : POINTER TO IoConfigConnector;
	NCOUNT : DINT;
END_VAR
END_METHOD

METHOD IODRVUPDATEMAPPING : UDINT
VAR_INPUT
	PTASKMAPLIST : POINTER TO IoConfigTaskMap;
	NCOUNT : DINT;
END_VAR
END_METHOD

METHOD IODRVWRITEPARAMETER : UDINT
VAR_INPUT
	PCONNECTOR : POINTER TO IoConfigConnector;
	PPARAMETER : POINTER TO IoConfigParameter;
	PDATA : POINTER TO BYTE;
	DWBITSIZE : DWORD;
	DWBITOFFSET : DWORD;
END_VAR
END_METHOD

METHOD QUERYINTERFACE : POINTER TO POINTER TO BYTE
VAR_INPUT
	IID : DWORD;
	PRESULT : POINTER TO UDINT;
END_VAR
END_METHOD

METHOD STATUSCHANGED : BOOL
END_METHOD

METHOD FB_EXIT : BOOL
VAR_INPUT
	BINCOPYCODE : BOOL;
END_VAR
END_METHOD

METHOD FB_INIT : BOOL
VAR_INPUT
	BINITRETAINS : BOOL;
	BINCOPYCODE : BOOL;
END_VAR
END_METHOD

METHOD EVENTCALLBACK : UDINT
VAR_INPUT
	PEVENTPARAM : POINTER TO EventParam;
END_VAR
END_METHOD

METHOD REGISTEREVENT
END_METHOD

METHOD UNREGISTEREVENT
END_METHOD

(* ---- L_MC1P_AXISEXTENSION_9400HL.fb ---- *)
FUNCTION_BLOCK L_MC1P_AXISEXTENSION_9400HL EXTENDS L_MC1P_AxisExtensionEmpty
VAR
	ECATCOMM : L_MC1P_CommECAT;
	CONFIGDRIVE : L_MC1P_Config_94HL_ETC;
	DRIVESCALING : L_MC1P_DriveScaling_94HL;
	DRIVESPECIFIC : L_MC1P_DriveSpecific_9400HL;
	FBEXTENDEDMAPPINGACCESS : L_MC1P_ExtendedMappingAccess;
	ITFCOMM : L_MC1P_ICommunication;
	ITFCONFIGDRIVE : L_MC1P_IConfigureDrive;
	ITFDRIVESCALING : L_MC1P_IDriveScaling;
	ITFDRIVESPECIFIC : L_MC1P_IDriveSpecificImplBase;
	ITFEXTENDEDMAPPINGACCESS : L_MC1P_IExtendedMappingAccess;
END_VAR
END_FUNCTION_BLOCK

(* ---- L_MC1P_AXISEXTENSION_9400HL_CAN.fb ---- *)
FUNCTION_BLOCK L_MC1P_AXISEXTENSION_9400HL_CAN EXTENDS L_MC1P_AxisExtensionEmpty
VAR
	CANCOMM : L_MC1P_CommCAN;
	CONFIGDRIVE : L_MC1P_Config_94HL_ETC;
	DRIVESCALING : L_MC1P_DriveScaling_94HL;
	DRIVESPECIFIC : L_MC1P_DriveSpecific_9400HL;
	FBEXTENDEDMAPPINGACCESS : L_MC1P_ExtendedMappingAccess;
	ITFCOMM : L_MC1P_ICommunication;
	ITFCONFIGDRIVE : L_MC1P_IConfigureDrive;
	ITFDRIVESCALING : L_MC1P_IDriveScaling;
	ITFDRIVESPECIFIC : L_MC1P_IDriveSpecificImplBase;
	ITFEXTENDEDMAPPINGACCESS : L_MC1P_IExtendedMappingAccess;
END_VAR
END_FUNCTION_BLOCK

(* ---- L_MC1P_AXISEXTENSION_ENCBPB.fb ---- *)
FUNCTION_BLOCK L_MC1P_AXISEXTENSION_ENCBPB EXTENDS L_MC1P_AxisExtensionEmpty
VAR
	DRIVESPECIFIC : L_MC1P_DriveSpecific_Enc_Bpb;
	DRIVESCALING : L_MC1P_DriveScaling;
	ITFDRIVESCALING : L_MC1P_IDriveScaling;
	ITFDRIVESPECIFIC : L_MC1P_IDriveSpecificImplBase;
END_VAR
END_FUNCTION_BLOCK

(* ---- L_MC1P_AXISEXTENSION_ENCFREE.fb ---- *)
FUNCTION_BLOCK L_MC1P_AXISEXTENSION_ENCFREE EXTENDS L_MC1P_AxisExtensionEmpty
VAR
	DRIVESPECIFIC : L_MC1P_DriveSpecific_Enc_Free;
	DRIVESCALING : L_MC1P_DriveScaling;
	ITFDRIVESCALING : L_MC1P_IDriveScaling;
	ITFDRIVESPECIFIC : L_MC1P_IDriveSpecificImplBase;
END_VAR
END_FUNCTION_BLOCK

(* ---- L_MC1P_AXISEXTENSION_ENCI500.fb ---- *)
FUNCTION_BLOCK L_MC1P_AXISEXTENSION_ENCI500 EXTENDS L_MC1P_AxisExtensionEmpty
VAR
	I500COMM : L_MC1P_CommECAT;
	DRIVESPECIFIC : L_MC1P_DriveSpecific_Enc_i500;
	DRIVESCALING : L_MC1P_DriveScaling;
	ITFCOMM : L_MC1P_ICommunication;
	ITFDRIVESCALING : L_MC1P_IDriveScaling;
	ITFDRIVESPECIFIC : L_MC1P_IDriveSpecificImplBase;
END_VAR
END_FUNCTION_BLOCK

(* ---- L_MC1P_AXISEXTENSION_ENCI900_ECAT.fb ---- *)
FUNCTION_BLOCK L_MC1P_AXISEXTENSION_ENCI900_ECAT EXTENDS L_MC1P_AxisExtensionEmpty
VAR
	CONFIGAXIS : L_MC1P_Config_i900_Enc_Drive;
	I900COMM : L_MC1P_CommECAT;
	FBEXTENDEDMAPPINGACCESS : L_MC1P_ExtendedMappingAccess;
	DRIVESPECIFIC : L_MC1P_DriveSpecific_Enc_i950 := STRUCT(xCheckCommunicationState := TRUE);
	DRIVESCALING : L_MC1P_DriveScaling_Enci900;
	ITFCOMM : L_MC1P_ICommunication;
	ITFCONFIGDRIVE : L_MC1P_IConfigureDrive;
	ITFDRIVESCALING : L_MC1P_IDriveScaling;
	ITFDRIVESPECIFIC : L_MC1P_IDriveSpecificImplBase;
	ITFEXTENDEDMAPPINGACCESS : L_MC1P_IExtendedMappingAccess;
END_VAR
END_FUNCTION_BLOCK

(* ---- L_MC1P_AXISEXTENSION_ENCI900_TARGET.fb ---- *)
FUNCTION_BLOCK L_MC1P_AXISEXTENSION_ENCI900_TARGET EXTENDS L_MC1P_AxisExtensionEmpty
VAR_INPUT
	COMM : L_MC1P_Commi900;
	CONFIG : L_MC1P_Config_i900_Enc_Drive;
END_VAR
VAR
	DRIVESPECIFIC : L_MC1P_DriveSpecific_Enc_i950;
	DRIVESCALING : L_MC1P_DriveScaling_Enci900;
	ITFCOMM : L_MC1P_ICommunication;
	ITFCONFIGDRIVE : L_MC1P_IConfigureDrive;
	ITFDRIVESCALING : L_MC1P_IDriveScaling;
	ITFDRIVESPECIFIC : L_MC1P_IDriveSpecificImplBase;
END_VAR
END_FUNCTION_BLOCK

(* ---- L_MC1P_AXISEXTENSION_ENCIOETC.fb ---- *)
FUNCTION_BLOCK L_MC1P_AXISEXTENSION_ENCIOETC EXTENDS L_MC1P_AxisExtensionEmpty
VAR
	DRIVESPECIFIC : L_MC1P_DriveSpecific_Enc_IOETC;
	DRIVESCALING : L_MC1P_DriveScaling;
	ITFDRIVESCALING : L_MC1P_IDriveScaling;
	ITFDRIVESPECIFIC : L_MC1P_IDriveSpecificImplBase;
END_VAR
END_FUNCTION_BLOCK

(* ---- L_MC1P_AXISEXTENSION_GENERICDRIVE.fb ---- *)
FUNCTION_BLOCK L_MC1P_AXISEXTENSION_GENERICDRIVE EXTENDS L_MC1P_AxisExtensionEmpty
VAR
	CONFIGDRIVE : L_MC1P_Config_GenericDrive;
	DRIVESCALING : L_MC1P_DriveScaling_GenericDrive;
	DRIVESPECIFIC : L_MC1P_DriveSpecific_Generic;
	ECATCOMM : L_MC1P_CommECAT;
	FBEXTENDEDMAPPINGACCESS : L_MC1P_ExtendedMappingAccess;
	GETTYPE : L_MC1P_AxisExtensionTypes;
	ITFCOMM : L_MC1P_ICommunication;
	ITFCONFIGDRIVE : L_MC1P_IConfigureDrive;
	ITFDRIVESCALING : L_MC1P_IDriveScaling;
	ITFDRIVESPECIFIC : L_MC1P_IDriveSpecificImplBase;
	ITFEXTENDEDMAPPINGACCESS : L_MC1P_IExtendedMappingAccess;
END_VAR
END_FUNCTION_BLOCK

METHOD SETBASICINITIALISATION
VAR_INPUT
	ITFGENERICCONFIG : L_MC1P_IGenericAxisConfiguration;
END_VAR
VAR_IN_OUT
	AXIS : _AXIS_REF_REAL;
END_VAR
END_METHOD

(* ---- L_MC1P_AXISEXTENSION_I500_CAN.fb ---- *)
FUNCTION_BLOCK L_MC1P_AXISEXTENSION_I500_CAN EXTENDS L_MC1P_AxisExtensionEmpty
VAR_INPUT
	DRIVESPECIFIC : L_MC1P_DriveSpecific_i500;
END_VAR
VAR
	CONFIGDRIVE : L_MC1P_Config_i500;
	DRIVESCALING : L_MC1P_DriveScaling_i500;
	CANCOMM : L_MC1P_CommCAN;
	ITFCOMM : L_MC1P_ICommunication;
	ITFCONFIGDRIVE : L_MC1P_IConfigureDrive;
	ITFDRIVESCALING : L_MC1P_IDriveScaling;
	ITFDRIVESPECIFIC : L_MC1P_IDriveSpecificImplBase;
END_VAR
END_FUNCTION_BLOCK

METHOD FB_INIT : BOOL
VAR_INPUT
	BINITRETAINS : BOOL;
	BINCOPYCODE : BOOL;
END_VAR
END_METHOD

(* ---- L_MC1P_AXISEXTENSION_I500_ECAT.fb ---- *)
FUNCTION_BLOCK L_MC1P_AXISEXTENSION_I500_ECAT EXTENDS L_MC1P_AxisExtensionEmpty
VAR_INPUT
	DRIVESPECIFIC : L_MC1P_DriveSpecific_i500;
END_VAR
VAR
	CONFIGDRIVE : L_MC1P_Config_i500;
	DRIVESCALING : L_MC1P_DriveScaling_i500;
	ECATCOMM : L_MC1P_CommECAT;
	FBEXTENDEDMAPPINGACCESS : L_MC1P_ExtendedMappingAccess;
	ITFCOMM : L_MC1P_ICommunication;
	ITFCONFIGDRIVE : L_MC1P_IConfigureDrive;
	ITFDRIVESCALING : L_MC1P_IDriveScaling;
	ITFDRIVESPECIFIC : L_MC1P_IDriveSpecificImplBase;
	ITFEXTENDEDMAPPINGACCESS : L_MC1P_IExtendedMappingAccess;
END_VAR
END_FUNCTION_BLOCK

(* ---- L_MC1P_AXISEXTENSION_I700.fb ---- *)
FUNCTION_BLOCK L_MC1P_AXISEXTENSION_I700 EXTENDS L_MC1P_AxisExtensionEmpty
VAR
	CONFIGDRIVE : L_MC1P_Config_i700_ETC;
	ECATCOMM : L_MC1P_CommECAT;
	FBEXTENDEDMAPPINGACCESS : L_MC1P_ExtendedMappingAccess;
	DRIVESCALING : L_MC1P_DriveScaling_i7xx;
	BRAKE : L_MC1P_BrakeControl;
	DRIVESPECIFIC : L_MC1P_DriveSpecific_i700;
	ITFCOMM : L_MC1P_ICommunication;
	ITFCONFIGDRIVE : L_MC1P_IConfigureDrive;
	ITFDRIVESCALING : L_MC1P_IDriveScaling;
	ITFDRIVESPECIFIC : L_MC1P_IDriveSpecificImplBase;
	ITFEXTENDEDMAPPINGACCESS : L_MC1P_IExtendedMappingAccess;
END_VAR
END_FUNCTION_BLOCK

METHOD FB_INIT : BOOL
VAR_INPUT
	BINITRETAINS : BOOL;
	BINCOPYCODE : BOOL;
END_VAR
END_METHOD

(* ---- L_MC1P_AXISEXTENSION_I750.fb ---- *)
FUNCTION_BLOCK L_MC1P_AXISEXTENSION_I750 EXTENDS L_MC1P_AxisExtensionEmpty
VAR
	CONFIGDRIVE : L_MC1P_Config_i900Adv_ETC;
	ECATCOMM : L_MC1P_CommECAT;
	FBEXTENDEDMAPPINGACCESS : L_MC1P_ExtendedMappingAccess;
	DRIVESCALING : L_MC1P_DriveScaling_i7xx;
	BRAKE : L_MC1P_BrakeControl;
	DRIVESPECIFIC : L_MC1P_DriveSpecific_i750;
	ITFCOMM : L_MC1P_ICommunication;
	ITFCONFIGDRIVE : L_MC1P_IConfigureDrive;
	ITFDRIVESCALING : L_MC1P_IDriveScaling;
	ITFDRIVESPECIFIC : L_MC1P_IDriveSpecificImplBase;
	ITFEXTENDEDMAPPINGACCESS : L_MC1P_IExtendedMappingAccess;
END_VAR
END_FUNCTION_BLOCK

METHOD FB_INIT : BOOL
VAR_INPUT
	BINITRETAINS : BOOL;
	BINCOPYCODE : BOOL;
END_VAR
END_METHOD

(* ---- L_MC1P_AXISEXTENSION_I950.fb ---- *)
FUNCTION_BLOCK L_MC1P_AXISEXTENSION_I950 EXTENDS L_MC1P_AxisExtensionEmpty
VAR
	CONFIGDRIVE : L_MC1P_Config_i900Adv_ETC := STRUCT(xCiA402Advanced := FALSE);
	ECATCOMM : L_MC1P_CommECAT;
	FBEXTENDEDMAPPINGACCESS : L_MC1P_ExtendedMappingAccess;
	BRAKE : L_MC1P_BrakeControl;
	DRIVESCALING : L_MC1P_DriveScaling_i7xx;
	DRIVESPECIFIC : L_MC1P_DriveSpecific_i950;
	ITFCOMM : L_MC1P_ICommunication;
	ITFCONFIGDRIVE : L_MC1P_IConfigureDrive;
	ITFDRIVESCALING : L_MC1P_IDriveScaling;
	ITFDRIVESPECIFIC : L_MC1P_IDriveSpecificImplBase;
	ITFEXTENDEDMAPPINGACCESS : L_MC1P_IExtendedMappingAccess;
END_VAR
END_FUNCTION_BLOCK

METHOD FB_INIT : BOOL
VAR_INPUT
	BINITRETAINS : BOOL;
	BINCOPYCODE : BOOL;
END_VAR
END_METHOD

(* ---- L_MC1P_AXISEXTENSION_I950_CIAADV.fb ---- *)
FUNCTION_BLOCK L_MC1P_AXISEXTENSION_I950_CIAADV EXTENDS L_MC1P_AxisExtensionEmpty
VAR
	CONFIGDRIVE : L_MC1P_Config_i900Adv_ETC := STRUCT(xCiA402Advanced := TRUE);
	ECATCOMM : L_MC1P_CommECAT;
	FBEXTENDEDMAPPINGACCESS : L_MC1P_ExtendedMappingAccess;
	DRIVESCALING : L_MC1P_DriveScaling_i7xx;
	BRAKE : L_MC1P_BrakeControl;
	DRIVESPECIFIC : L_MC1P_DriveSpecific_i950Adv;
	ITFCOMM : L_MC1P_ICommunication;
	ITFCONFIGDRIVE : L_MC1P_IConfigureDrive;
	ITFDRIVESCALING : L_MC1P_IDriveScaling;
	ITFDRIVESPECIFIC : L_MC1P_IDriveSpecificImplBase;
	ITFEXTENDEDMAPPINGACCESS : L_MC1P_IExtendedMappingAccess;
END_VAR
END_FUNCTION_BLOCK

METHOD FB_INIT : BOOL
VAR_INPUT
	BINITRETAINS : BOOL;
	BINCOPYCODE : BOOL;
END_VAR
END_METHOD

(* ---- L_MC1P_AXISEXTENSION_I950_DRIVE.fb ---- *)
FUNCTION_BLOCK L_MC1P_AXISEXTENSION_I950_DRIVE EXTENDS L_MC1P_AxisExtensionEmpty
VAR_INPUT
	CONFIGDRIVE : L_MC1P_Config_i900_Drive;
	COMM : L_MC1P_Commi900;
END_VAR
VAR
	DRIVESCALING : L_MC1P_DriveScaling_i7xx;
	BRAKE : L_MC1P_BrakeControlBase;
	DRIVESPECIFIC : L_MC1P_DriveSpecific_i950_Drive;
	ITFCOMM : L_MC1P_ICommunication;
	ITFCONFIGDRIVE : L_MC1P_IConfigureDrive;
	ITFDRIVESCALING : L_MC1P_IDriveScaling;
	ITFDRIVESPECIFIC : L_MC1P_IDriveSpecificImplBase;
END_VAR
END_FUNCTION_BLOCK

METHOD FB_INIT : BOOL
VAR_INPUT
	BINITRETAINS : BOOL;
	BINCOPYCODE : BOOL;
END_VAR
END_METHOD

(* ---- L_MC1P_AXISEXTENSIONEMPTY.fb ---- *)
FUNCTION_BLOCK L_MC1P_AXISEXTENSIONEMPTY
VAR
	GETTYPE : L_MC1P_AxisExtensionTypes;
	ITFCOMM : L_MC1P_ICommunication;
	ITFCONFIGDRIVE : L_MC1P_IConfigureDrive;
	ITFDRIVESCALING : L_MC1P_IDriveScaling;
	ITFDRIVESPECIFIC : L_MC1P_IDriveSpecificImplBase;
	ITFEXTENDEDMAPPINGACCESS : L_MC1P_IExtendedMappingAccess;
END_VAR
END_FUNCTION_BLOCK

METHOD SETBASICINITIALISATION
VAR_INPUT
	ITFGENERICCONFIG : L_MC1P_IGenericAxisConfiguration;
END_VAR
VAR_IN_OUT
	AXIS : _AXIS_REF_REAL;
END_VAR
END_METHOD

METHOD FB_EXIT : BOOL
VAR_INPUT
	BINCOPYCODE : BOOL;
END_VAR
END_METHOD

(* ---- L_MC1P_AXISINTERFACE.fb ---- *)
FUNCTION_BLOCK L_MC1P_AXISINTERFACE EXTENDS L_MC1P_Template
VAR_INPUT
	XENABLE : BOOL;
	EXTCONTROLLER : L_MC1P_IControllerInterface;
END_VAR
VAR_OUTPUT
	XVALID : BOOL;
	XBUSY : BOOL;
	XERROR : BOOL;
	EERRORID : L_IE1P_Error;
END_VAR
VAR
	XENABLEOLD : BOOL;
END_VAR
END_FUNCTION_BLOCK

(* ---- L_MC1P_AXISMANAGEMENTFUNCTION.fb ---- *)
FUNCTION_BLOCK L_MC1P_AXISMANAGEMENTFUNCTION
VAR
	LMAXISMANAGEMENTFUNCTION : ARRAY [1..L_MC1P_Constants.gc_MaxAxisCount] OF L_MC1P_IManagementFunction;
	DIAXISCOUNT : DINT;
END_VAR
END_FUNCTION_BLOCK

METHOD FINDAXISBYNAME : POINTER TO AXIS_REF
VAR_IN_OUT
	SAXISNAME : STRING;
END_VAR
END_METHOD

METHOD GETFIRSTAXIS : POINTER TO AXIS_REF
VAR_INPUT
	PIDX : POINTER TO DINT;
END_VAR
END_METHOD

METHOD GETNEXTAXIS : POINTER TO AXIS_REF
VAR_INPUT
	PIDX : POINTER TO DINT;
END_VAR
END_METHOD

METHOD REGISTERAXIS : BOOL
VAR_INPUT
	ITFMANAGE : L_MC1P_IManagementFunction;
END_VAR
END_METHOD

(* ---- L_MC1P_AXISMASTERVALUESEMPTY.fb ---- *)
FUNCTION_BLOCK L_MC1P_AXISMASTERVALUESEMPTY
VAR
	FBSTEADYSTATE : L_MC1P_SteadyState;
	ACTACCELERATION : LREAL;
	ACTPOSITION : LREAL;
	ACTTORQUE : LREAL;
	ACTVELOCITY : LREAL;
	CYCLELENGTH : LREAL;
	FEEDCONSTANT : LREAL;
	GETMASTERID : POINTER TO BYTE;
	SETACCELERATIONFORSYNC : LREAL;
	SETPOSITIONFORSYNC : LREAL;
	SETTORQUEFORSYNC : LREAL;
	SETVELOCITYFORSYNC : LREAL;
	TASKCYCLE : LREAL;
	TRAVERSINGRANGE : L_MC1P_TraversingRange;
END_VAR
END_FUNCTION_BLOCK

METHOD GETDIRECTION : WORD
VAR_INPUT
	VALUESOURCE : MC_SOURCE;
END_VAR
END_METHOD

METHOD GETMASTERERROR : BOOL
VAR_OUTPUT
	EERRORID : L_IE1P_Error;
END_VAR
END_METHOD

METHOD GETSTEADYSTATE : POINTER TO L_MC1P_SteadyState
END_METHOD

(* ---- L_MC1P_AXISRETAINMANGAEMENT.fb ---- *)
FUNCTION_BLOCK L_MC1P_AXISRETAINMANGAEMENT
VAR_OUTPUT
	XERROR : BOOL;
END_VAR
VAR
	XINIT : BOOL := FALSE;
	ERRORHANDLE : SysTypes.RTS_IEC_HANDLE := 0;
	MODULEHANDLE : SysTypes.RTS_IEC_HANDLE := 0;
	DWLENGTH : DWORD;
	XMEMVALID : BOOL := FALSE;
	PSTARTADRESS : POINTER TO DWORD;
	PMEMADRESS : POINTER TO DWORD;
	PMEMADRESSMIRROR : POINTER TO DWORD;
	DWMEMSIZE : DWORD;
	DIAXISCOUNT : DINT := 0;
	LMAXISINFORMATION : ARRAY [1..L_MC1P_Constants.gc_MaxRetainAxis] OF L_MC1P_AxisRetainInformation;
	WSTEP : WORD := 0;
	XCONFIGCHANGED : BOOL;
	DATAMEMORYAREA : L_SSYP_PersistantDataMemoryArea;
	DWVERSION : DWORD;
	XINITIALAREA : BOOL := FALSE;
	DWTOTALSIZE1 : DWORD;
	DWTOTALSIZE2 : DWORD;
	PADWDUMMY1 : POINTER TO ARRAY [1..100] OF DWORD;
	PADWDUMMY2 : POINTER TO ARRAY [1..100] OF DWORD;
	WINTSTATE : WORD;
	DIIDX : DINT;
	BYMEMVERSION : BYTE;
	SINSTANCESTRFULL : STRING(255);
	BYACTMEMVERSION : BYTE := 2;
END_VAR
END_FUNCTION_BLOCK

METHOD CHECKMEMORY
END_METHOD

METHOD GETDATA : BOOL
VAR_IN_OUT
	AXISRETAIN : L_MC1P_AxisRetainInformation;
END_VAR
END_METHOD

METHOD READDWORD : DWORD
VAR_IN_OUT
	DWSIZEREAD : DWORD;
END_VAR
END_METHOD

METHOD READMEMORY
END_METHOD

METHOD REINITMEMORY
VAR_INPUT
	PDATA : POINTER TO DWORD;
	XMIRROR : BOOL;
END_VAR
END_METHOD

METHOD SEARCHDATA : BOOL
VAR_IN_OUT
	DWSIZEREAD : DWORD;
	AXISRETAIN : L_MC1P_AxisRetainInformation;
END_VAR
END_METHOD

METHOD SETACTIVEMEMAREA
VAR_INPUT
	XMIRROR : BOOL;
END_VAR
END_METHOD

METHOD SETMEMORYINVALID
END_METHOD

METHOD WRITEAXISDATA
END_METHOD

METHOD WRITEDWORD : DWORD
VAR_INPUT
	PMEMBASE : POINTER TO DWORD;
	DWDATA : DWORD;
END_VAR
VAR_IN_OUT
	DWSIZEWRITE : DWORD;
END_VAR
END_METHOD

METHOD FB_EXIT : BOOL
VAR_INPUT
	BINCOPYCODE : BOOL;
END_VAR
END_METHOD

METHOD FB_INIT : BOOL
VAR_INPUT
	BINITRETAINS : BOOL;
	BINCOPYCODE : BOOL;
END_VAR
END_METHOD

METHOD REGISTERAXIS
VAR_INPUT
	AXISGUID : L_MC1P_AxisGUID;
END_VAR
END_METHOD

METHOD REGISTERAXIS2 : POINTER TO L_MC1P_AxisRetainInformation
VAR_INPUT
	AXISGUID : L_MC1P_AxisGUID;
	ITFRETAIN : L_MC1P_IRetainFunction;
END_VAR
END_METHOD

METHOD INITMEMFORAXIS
VAR_INPUT
	PDATA : POINTER TO DWORD;
	XMIRROR : BOOL;
END_VAR
VAR_IN_OUT
	DWWRITEOFFSET : DWORD;
	AXISRETAININFORMATION : L_MC1P_AxisRetainInformation;
END_VAR
END_METHOD

METHOD WRITEADDSIZE
VAR_INPUT
	PDATA : POINTER TO DWORD;
	DWADDSIZE : DWORD;
END_VAR
END_METHOD

METHOD WRITEHEADER
VAR_INPUT
	PDATA : POINTER TO DWORD;
END_VAR
END_METHOD

(* ---- L_MC1P_AXISSIMREADPRM.fb ---- *)
FUNCTION_BLOCK L_MC1P_AXISSIMREADPRM EXTENDS L_UBUP_FreeRunTask
VAR_INPUT
	UIDEVICEID : UINT;
	PPARAMDATA : POINTER TO L_MC1P_ParameterDataSim;
	WPARAMCOUNT : WORD;
	PPARAMDATAIGNORE : POINTER TO L_MC1P_ParameterDataSim;
	WPARAMCOUNTIGNORE : WORD;
END_VAR
VAR
	PARSIMWRITE : L_MC1P_ParSimWrite;
	SBASEPATH : STRING(255);
END_VAR
END_FUNCTION_BLOCK

METHOD CUSTOMIZEERRORCODE : L_IE1P_Error
VAR_INPUT
	IERRORID : INT;
END_VAR
END_METHOD

METHOD EXECUTEIMPL : UDINT
END_METHOD

METHOD FB_INIT : BOOL
VAR_INPUT
	BINITRETAINS : BOOL;
	BINCOPYCODE : BOOL;
END_VAR
END_METHOD

(* ---- L_MC1P_AXISSIMULATION.fb ---- *)
FUNCTION_BLOCK L_MC1P_AXISSIMULATION
VAR_INPUT
	SCIODATA : L_MC1P_AxisSimIOData;
	SCPARMECHANIC : L_MC1P_ParMechanic;
	SCPAROBDDRIVE : L_MC1P_AxisSimulationSdoData;
	SCPARGENERAL : L_MC1P_ParGeneralMechanic;
	LRINITIALPOSITION : LREAL;
	EINITOBDDRIVEMODE : UINT := 0;
END_VAR
VAR_OUTPUT
	XBUSY : BOOL;
END_VAR
VAR
	COMMUNICATION : L_MC1P_CommSim;
	APARAMDATA : ARRAY [1..c_MaxSimData] OF L_MC1P_ParameterDataSim;
	APRMIGNOREDATA : ARRAY [1..c_MaxPrmIgnoreData] OF L_MC1P_ParameterDataSim;
	TRANSMITDATA : L_MC1P_AxisSimulationPDOdataToDrive;
	RECIEVEDATA : L_MC1P_AxisSimulationPDOdataFromDrive;
	LWTRANSDATA : LWORD;
	LWTRANSDATASAVE : LWORD;
	WTRANSELEMENTS : WORD;
	ATRANSELEMENT : ARRAY [1..c_wMaxTransElem] OF L_MC1P_MappedElement;
	ATRANSELEMENTADRESS : ARRAY [1..L_MC1P_Constants.gc_Trans_MaxDataIndex] OF POINTER TO L_MC1P_MappedElement;
	ATRANSELEMENTADRESSSAVE : ARRAY [1..L_MC1P_Constants.gc_Trans_MaxDataIndex] OF POINTER TO L_MC1P_MappedElement;
	LWRECDATA : LWORD;
	LWRECDATASAVE : LWORD;
	WRECEIVEELEMENTS : WORD;
	ARECEIVEELEMENT : ARRAY [1..c_wMaxRecElem] OF L_MC1P_MappedElement;
	ARECEIVEELEMENTADRESS : ARRAY [1..L_MC1P_Constants.gc_Rec_MaxDataIndex] OF POINTER TO L_MC1P_MappedElement;
	ARECEIVEELEMENTADRESSSAVE : ARRAY [1..L_MC1P_Constants.gc_Rec_MaxDataIndex] OF POINTER TO L_MC1P_MappedElement;
	IBUSDEADCYCLES : INT := 2;
	IINDEXPDO : INT := 1;
	ASCPDO_P2D : ARRAY [0..(ciPDO_BufferSize - 1)] OF L_MC1P_AxisSimulationPDOdataToDrive;
	ASCPDO_D2P : ARRAY [0..(ciPDO_BufferSize - 1)] OF L_MC1P_AxisSimulationPDOdataFromDrive;
	SYSTEMSIMULATION : L_MC1P_SimMotorCtrl;
	MECHANICSIMULATION : L_MC1P_SimMechanic;
	ITFMECHANICMODELDEFAULT : L_MC1P_IMechanicSimulation := MechanicSimulation;
	ITFMECHANICMODELACT : L_MC1P_IMechanicSimulation := itfMechanicModelDefault;
	TRANSMITDATASCALED : L_MC1P_AxisSimulationPDOdataToDriveScaled;
	RECIEVEDATASCALED : L_MC1P_AxisSimulationPDOdataFromDriveScaled;
	XREADPARSET : BOOL;
	AXISSIMREADPRM : L_MC1P_AxisSimReadPRM;
	XGENERRORREAKTINDEVICESAVE : BOOL;
	C_WMAXTRANSELEM : WORD := 20;
	C_WMAXRECELEM : WORD := 38;
	C_MAXSIMDATA : WORD := 90;
	C_MAXPRMIGNOREDATA : WORD := 5;
	CIPDO_BUFFERSIZE : INT := 10;
	COMMSIMULATION : L_MC1P_ICommmunicationSimulation;
	GETRECIEVEDATACONFIG : LWORD;
	GETTRANSMITDATACONFIG : LWORD;
	LOADFDB : LREAL;
	RECIEVEELEMCOUNT : WORD;
	RECIEVEELEMENT : POINTER TO L_MC1P_MappedElement;
	RECIEVEELEMENTADRESS : POINTER TO ARRAY [1..L_MC1P_Constants.gc_Rec_MaxDataIndex] OF POINTER TO L_MC1P_MappedElement;
	TRANSELEMCOUNT : WORD;
	TRANSELEMENT : POINTER TO L_MC1P_MappedElement;
	TRANSELEMENTADRESS : POINTER TO ARRAY [1..L_MC1P_Constants.gc_Trans_MaxDataIndex] OF POINTER TO L_MC1P_MappedElement;
END_VAR
END_FUNCTION_BLOCK

METHOD SETMECHANICMODEL : BOOL
VAR_INPUT
	ITFMECHANICMODEL : L_MC1P_IMechanicSimulation;
END_VAR
END_METHOD

METHOD CALCOPTIMIZEDMAPPINGINFO : BOOL
END_METHOD

METHOD GETBITNBR : WORD
VAR_INPUT
	LWMASK : LWORD;
END_VAR
END_METHOD

METHOD INITOBD : BOOL
END_METHOD

METHOD SETDRIVEDEPENDENTMAPPING : BOOL
VAR_IN_OUT
	AXIS : _AXIS_REF_REAL;
END_VAR
END_METHOD

METHOD SETPARAMETERINFO : BOOL
VAR_INPUT
	PARAMDATAIDX : WORD;
	WINDEX : WORD;
	BYSUBINDEX : BYTE;
	PDOMAPNBR : LWORD;
	PDATA : POINTER TO BYTE;
	BYNROFBYTE : BYTE;
	XSUPPORTED : BOOL;
	XWRITEACCESS : BOOL;
	XAXISOFFSET : BOOL;
	EFIXTOLREAL : L_MC1P_ScaleFixToLREAL := L_MC1P_ScaleFixToLREAL.None;
END_VAR
END_METHOD

METHOD FB_INIT : BOOL
VAR_INPUT
	BINITRETAINS : BOOL;
	BINCOPYCODE : BOOL;
END_VAR
END_METHOD

METHOD GETBUSVALUESP2D
VAR_IN_OUT
	AXIS : _AXIS_REF_REAL;
END_VAR
END_METHOD

METHOD WRITEBUSVALUESD2P
VAR_IN_OUT
	AXIS : _AXIS_REF_REAL;
END_VAR
END_METHOD

METHOD ACTIVATESIMULATION
VAR_IN_OUT
	AXIS : _AXIS_REF_REAL;
END_VAR
END_METHOD

METHOD CALCULATEINPUTDATA
VAR_IN_OUT
	AXIS : _AXIS_REF_REAL;
END_VAR
END_METHOD

METHOD CALCULATEOUTPUTDATA
VAR_IN_OUT
	AXIS : _AXIS_REF_REAL;
END_VAR
END_METHOD

METHOD DISABLESIMULATION
VAR_IN_OUT
	AXIS : _AXIS_REF_REAL;
END_VAR
END_METHOD

(* ---- L_MC1P_BASICACTUATINGSPEED.fb ---- *)
FUNCTION_BLOCK L_MC1P_BASICACTUATINGSPEED EXTENDS L_MC1P_Template
VAR_INPUT
	XENABLEINTERNALCONTROL : BOOL := FALSE;
	XREGULATORON : BOOL := FALSE;
	XRESETERROR : BOOL := FALSE;
	XSETDRIVEQSP : BOOL := FALSE;
	XENABLESETVEL : BOOL := FALSE;
	XINVERTDIRECTION : BOOL := FALSE;
	LRSETVEL : LREAL := 0.0;
	LRSETACC : LREAL := 0.0;
	LRSETDEC : LREAL := 0.0;
END_VAR
VAR_OUTPUT
	XINTERNALCONTROLACTIVE : BOOL;
	XBUSY : BOOL;
	XERROR : BOOL;
	EERRORID : L_IE1P_Error;
	XCOMMUNICATIONOK : BOOL;
	XAXISREADY : BOOL;
	XAXISENABLED : BOOL;
	XDRIVEWARNING : BOOL;
	XDRIVEERROR : BOOL;
	DWDRIVEERRORID : DWORD;
	XDRIVEQSPACTIVE : BOOL;
	LRACTVEL : LREAL;
	XDIRECTIONPOSITIVE : BOOL;
	XDIRECTIONNEGATIVE : BOOL;
	WDIGITALINPUTS : WORD;
END_VAR
VAR
	XINTERNALCONTROLVISU : BOOL;
	XREGULATORON_INT : BOOL := FALSE;
	XSETDRIVEQSP_INT : BOOL := FALSE;
	XRESETERROR_INT : BOOL := FALSE;
	XENABLESETVEL_INT : BOOL := FALSE;
	XINVERTDIRECTION_INT : BOOL := FALSE;
	LRSETVEL_INT : LREAL := 0.0;
	LRSETACC_INT : LREAL := 0.0;
	LRSETDEC_INT : LREAL := 0.0;
	LRSETACCOLD : LREAL := 0.0;
	LRSETDECOLD : LREAL := 0.0;
	LRSCALERPMTOUNITOLD : LREAL := 0.0;
	READAXISERROR : L_MC1P_ReadAxisError_Internal;
	FBRESET : L_MC1P_Reset_Internal;
	DWDIGIN : DWORD;
	PREALAXIS : POINTER TO _AXIS_REF_REAL;
	PWDUMMY : POINTER TO WORD;
	PXDUMMY : POINTER TO BOOL;
	BYSDORETRYCOUNTER : BYTE;
	XWAITFORPARAMETERWRITEDONE : BOOL;
	WRITEPARAMETER : L_DCO_WriteDriveParameter;
	WSTEP : WORD;
	DWDELTASPEED : DWORD;
	WDELTATIME : WORD;
	XINTERNALCONTROLACTIVEOLD : BOOL;
	WLCONTROLWORD : WORD;
	WLCONTROLWORD2 : WORD;
	WLCONTROLWORD3 : WORD;
	WLCONTROLWORD4 : WORD;
	WLSTATUSWORD : WORD;
	WLSTATUSWORD2 : WORD;
	PITFMANIPULATEACTVALUES : POINTER TO L_Mc1P_IManipulateActValues;
	MAX_SDO_RETRIES : WORD := 3;
	LCONTROLWORD : WORD;
	LCONTROLWORD2 : WORD;
	LCONTROLWORD3 : WORD;
	LCONTROLWORD4 : WORD;
	LSTATUSWORD : WORD;
	LSTATUSWORD2 : WORD;
END_VAR
END_FUNCTION_BLOCK

METHOD CALCACCVALUES
VAR_INPUT
	LRACC : LREAL;
END_VAR
VAR_OUTPUT
	DWDELTASPEED : DWORD;
	WDELTATIME : WORD;
END_VAR
VAR_IN_OUT
	REALAXIS : _AXIS_REF_REAL;
END_VAR
END_METHOD

METHOD CHECKACCDECCHANGED
VAR_IN_OUT
	REALAXIS : _AXIS_REF_REAL;
END_VAR
END_METHOD

METHOD MANIPULATEACTVALUES
VAR_IN_OUT
	AXIS : AXIS_REF;
END_VAR
END_METHOD

(* ---- L_MC1P_BRAKECONTROL.fb ---- *)
FUNCTION_BLOCK L_MC1P_BRAKECONTROL EXTENDS L_MC1P_BrakeControlBase
VAR_INPUT
	LRTORQUEADD : LREAL;
	XSTARTINGTORQUE2 : BOOL;
	LRBRAKERAMPTIME : REFERENCE TO LREAL;
	XBRAKEACCDEPENDING : REFERENCE TO BOOL;
	LRSPEEDMIN : LREAL;
	LRRAMPWATCHTIME : LREAL;
	WSOURCESTARTVALUE : REFERENCE TO WORD;
	ALRMSTARTVALUE : REFERENCE TO ARRAY [1..2] OF LREAL;
	LREFFECTIVESTARTINGTORQUE : REFERENCE TO LREAL;
END_VAR
VAR
	LRSPEEDSET : LREAL;
	LRSPEEDACT : LREAL;
	XMOTORPHASESOK : BOOL := TRUE;
	MCTRLCONF : L_MC1P_MctrlControl := L_MC1P_MctrlControl.mcStandard;
	XESSACTIVE : BOOL := FALSE;
	XFLYINGSYNCBUSY : BOOL;
	XDCBRAKEISACTIVE : BOOL := FALSE;
	XDCBRAKEINSTEADQSP : BOOL := FALSE;
	XQSPISACTIVE : BOOL := FALSE;
	XSLIPCTRLACTIVE : BOOL := FALSE;
	XMAGNETISATIONISFINISHED : BOOL := FALSE;
	XUVDETECTED : BOOL;
	LRMAGNETISATIONTIME : LREAL := 1.0;
	LRTASKCYCLE : LREAL := 0.001;
	LRREFERENCETORQUE : LREAL;
	XINVERTBRAKECTRL : BOOL;
	XBRAKESTATEINPUT : BOOL;
	XIMPBRAKEREACTION : BOOL;
	LRBRAKEOBSERVATIONDELAY : LREAL;
	XBRAKEFEEDBACK : BOOL;
	XGETCINH_NOBRAKE : BOOL;
	XBRKSETCINH : BOOL;
	LRSETSPEEDOUT : LREAL;
	XBRAKEAPPLIED : BOOL;
	LRTORQUESET : LREAL;
	LRSPEEDSETOLD : LREAL;
	LRSPEEDACTOLD : LREAL;
	LRSPEEDCTRLINTVALUESET : LREAL;
	XLASTSPEEDBELOWMINSPEED : BOOL;
	LRTIMEOUTCOUNTER : LREAL;
	LRRELEASECOUNTER : LREAL;
	LROBSERVATIONCOUNTER : LREAL;
	XAUTOSUPERVISOROLD : BOOL;
	LRTORQUEACTFILTERED : LREAL;
	XSPEEDEQZERO : BOOL;
	XAXISERROR : BOOL;
	XQSPACTIVE : BOOL;
	XSETSPEEDTOZERO : BOOL;
	XAXISCINH : BOOL;
	LRAXISDECERRSTOP : LREAL;
	LRAXISJERKERRSTOP : LREAL;
	XBRAKEMODEINIT : BOOL;
	LRDRIVEMODEOBERSERVATIONCOUNTER : LREAL;
	XCIASTATUS : BOOL;
	DIPOSACT2NDSOURCE : DINT;
	DIBRAKEPOSITION2NDSOURCE : DINT;
	X2NDPOSVALID : BOOL;
	READPOS2NDSOURCE : L_DCO_ReadDriveParameter;
	XACTIVATEBRAKEMODEOBSERVATION : BOOL := TRUE;
	XDELAYOPERATIONENABLEDINACTIVE : BOOL := TRUE;
	XCLOSEBRAKEBECAUSOFFAULTREACTION : BOOL := FALSE;
	XCLOSEBRAKEATQSPRAMPEND : BOOL := FALSE;
	BRAKELOGICINPLCACTIVE : BOOL;
	PINSTANCE : POINTER TO L_MC1P_BrakeControlBase;
	TORQUEPRECONTROLACTIVE : BOOL;
END_VAR
END_FUNCTION_BLOCK

METHOD BF_BRAKE
END_METHOD

METHOD CONNECTPARAMETER : BOOL
VAR_INPUT
	PBRAKEPARA : POINTER TO L_MC1P_BrakePara;
END_VAR
END_METHOD

METHOD INIT
VAR_INPUT
	WBRAKEMODEINDEXOFDRIVE : WORD;
	BYSUBINDEX : BYTE;
	SZSIZE : BYTE;
	DEFAULTVALUE : DWORD;
END_VAR
VAR_IN_OUT
	AXIS : AXIS_REF;
END_VAR
END_METHOD

METHOD SUPPORTEDFUNCTION : INT
END_METHOD

METHOD FB_INIT : BOOL
VAR_INPUT
	BINITRETAINS : BOOL;
	BINCOPYCODE : BOOL;
END_VAR
END_METHOD

METHOD MODEAUTOENTERBRAKECLOSED
END_METHOD

METHOD MODEAUTOSTATEBRAKECLOSED
END_METHOD

METHOD MODEAUTOENTERCLOSINGBRAKE
END_METHOD

METHOD MODEAUTOENTERRAMPDOWN
END_METHOD

METHOD MODEAUTOSTATECLOSINGBRAKE
END_METHOD

METHOD MODEAUTOSTATERAMPDOWN
END_METHOD

METHOD BRAKECLEARERROR
VAR_INPUT
	ERRORCODE : L_MC1P_BrakeErrorCodes;
END_VAR
END_METHOD

METHOD BRAKERAISEERROR
VAR_INPUT
	ERRORCODE : L_MC1P_BrakeErrorCodes;
END_VAR
END_METHOD

METHOD ACTSPEEDISBELOWMINSPEED : BOOL
END_METHOD

METHOD BF_BRAKECLOSE
END_METHOD

METHOD BF_BRAKEDIRECTMODE
VAR_INPUT
	XSETDIRECTMODE : BOOL;
END_VAR
END_METHOD

METHOD BF_BRAKEGETSTATE : L_MC1P_BrakeState
VAR_OUTPUT
	ESTATEOPERATION : INT;
END_VAR
END_METHOD

METHOD BF_BRAKEGETSTATE_STATECONTROL : L_MC1P_BrakeState
END_METHOD

METHOD BF_BRAKEOPEN
END_METHOD

METHOD BF_BRAKEOUTPUTS
END_METHOD

METHOD BF_FQSPACTIVE : BOOL
END_METHOD

METHOD BF_TRIPACTIVE : BOOL
END_METHOD

METHOD BRAKEMODEOFF
END_METHOD

METHOD BRAKEMODEVALID : BOOL
VAR_INPUT
	BRAKEMODE : L_MC1P_BrakeMode;
END_VAR
END_METHOD

METHOD CONVERTBRAKEMODE : L_MC1P_InternalBrakeMode
VAR_INPUT
	EMODE : L_MC1P_BrakeMode;
END_VAR
END_METHOD

METHOD GETACTSPEEDISBELOWMINSPEED : BOOL
END_METHOD

METHOD INITTORQUEPRECONTROL
END_METHOD

METHOD ISBRAKECLOSEREQUESTED : BOOL
END_METHOD

METHOD ISBRAKERELEASEREQUESTED : BOOL
END_METHOD

METHOD ISNOFEEDBACK : BOOL
END_METHOD

METHOD ISNOIMPBECAUSEOFDCBRAKE : BOOL
END_METHOD

METHOD MODEAUTO
END_METHOD

METHOD MODEAUTOSTATESUPERVISOR
END_METHOD

METHOD MODEDIRECTCONTROL
END_METHOD

METHOD MODEMANUAL
END_METHOD

METHOD RESETOUTPUTSTATE
END_METHOD

METHOD SETSPEEDISBELOWMINSPEED : BOOL
END_METHOD

METHOD SPEEDEQ0 : BOOL
VAR_INPUT
	LRACTSPEED : LREAL;
	LRACTSPEEDOLD : LREAL;
END_VAR
END_METHOD

METHOD GETACTVALUES
END_METHOD

METHOD SWITCHONCONTROL
VAR_INPUT
	XSWITCHONREQUEST : BOOL;
END_VAR
VAR_OUTPUT
	XSWITCHON : BOOL;
END_VAR
VAR_IN_OUT
	AXIS : AXIS_REF;
END_VAR
END_METHOD

METHOD SWITCHEDONSTATUS
VAR_INPUT
	XSWITCHEDONREQUEST : BOOL;
END_VAR
VAR_OUTPUT
	XSWITCHEDON : BOOL;
END_VAR
VAR_IN_OUT
	AXIS : AXIS_REF;
END_VAR
END_METHOD

METHOD MODEAUTOENTERIDLE
END_METHOD

METHOD MODEAUTOSTATEIDLE
END_METHOD

METHOD BRAKEPRECONTROLWHILECLOSING
END_METHOD

METHOD BRAKETORQUECONTROL : BOOL
END_METHOD

METHOD GENERATETORQUEPRECONTROL
VAR_INPUT
	PLRACTVAL : POINTER TO LREAL;
	LRENDVAL : LREAL;
END_VAR
END_METHOD

METHOD MODEAUTOENTERRELEASINGBRAKE
END_METHOD

METHOD MODEAUTOSTATERELEASINGBRAKE
END_METHOD
